(* IEC 61131-3 sources: plc_agent/plc_agent/data/rag_data/st/st_case_code, 701 files *)

(* ---- ACOSH.st ---- *)
FUNCTION ACOSH : REAL
VAR_INPUT
    X : REAL;
END_VAR
ACOSH := LN(SQRT(X * X - 1.0) + X);

(* revision history
hm		12 jan 2007	rev 1.0
	original version

hm		2. dec 2007	rev 1.1
	changed code for better performance

hm	16. mar. 2007		rev 1.2
	changed sequence of calculations to improve performance

hm	10. mar. 2009		rev 1.3
	real constants updated to new systax using dot

*)
END_FUNCTION

(* ---- ACOTH.st ---- *)
FUNCTION ACOTH : REAL
VAR_INPUT
    X : REAL;
END_VAR
ACOTH := LN((x+1.0)/(x-1.0))*0.5;

(* revision history
hm		12 jan 2007	rev 1.0
	original version

hm		5. jan 2008	rev 1.1
	improved code for better performance

hm	10. mar. 2009		rev 1.2
	real constants updated to new systax using dot

*)
END_FUNCTION

(* ---- AGDF.st ---- *)
FUNCTION AGDF : REAL
VAR_INPUT
    X : REAL;
END_VAR
AGDF := LN((1.0 + SIN(X)) / COS(X));

(* comment
the current implementation gives sufficient accuracy only up to X = 1.57 or an output > 10.
is X closer to PI/2 then the function is more and more unreliable
*)

(* revision history
hm	27. apr. 2008	rev 1.0
	original version

hm	10. mar. 2009	rev 1.1
	real constants updated to new systax using dot

*)
END_FUNCTION

(* ---- AIN.st ---- *)
FUNCTION AIN : REAL
VAR_INPUT
    in : DWORD;
    Bits : BYTE;
    sign : BYTE := 255;
    low : REAL;
    high : REAL := 10.0;
END_VAR

VAR_CONSTANT
    ff : DWORD := 16#FFFFFFFF;
END_VAR

VAR
    temp1 : DWORD;
    temp2 : DWORD;
    sx : BOOL;
END_VAR
(* extract the sign bit *)
IF sign < 32 THEN
	temp1 := SHR(in,sign);
	sx := temp1.0;
ELSE
	sx := FALSE;
END_IF;
temp1 := SHR(ff, 32-bits);
temp2 := in AND temp1;
AIN := (high - low) * DWORD_TO_REAL(temp2) / DWORD_TO_REAL(temp1) + low;
IF sx THEN AIN := -AIN; END_IF;

(* revision history
hm 18.8.2006	rev 1.1
	fixed an error with low value negative and high value 0.

hm 19.1.2007	rev 1.2
	fixed an error with sign bit.

hm	13.9.2007	rev 1.3
	changed code to avoid warning under codesys 2.8.1

hm	2. dec 2007	rev 1.4
	changed code for better performance

hm	16. mar 2008	rev 1.5
	added type conversions to avoid warnings under codesys 30
*)
END_FUNCTION

(* ---- AIR_DENSITY.st ---- *)
FUNCTION AIR_DENSITY : REAL
VAR_INPUT
    T : REAL;     // Temperature
    P : REAL;     // Pressure
    RH : REAL;    // Relative Humidity
END_VAR

VAR CONSTANT
    RL : REAL := 287.05;   // Constant value for RL
    RX : REAL := 0.003773319;  // Constant value for RX
END_VAR
AIR_DENSITY := OSCAT_BASIC.phys.PN * (1.0 - RH * SDD(T, TRUE) * RX / P) / (RL * ( T - OSCAT_BASIC.phys.T0));

(* original code used for rev 1.0

SDD := SDD(T,FALSE);
RF := RL / (1- RH*SDD/P*RX);
Air_density := P / (RF * (T-TK));

*)

(* revision history

hm	29.10.2007	rev 1.0
	original version

hm	4.12.2007		rev 1.1
	changed code for better performance

hm	18. oct. 2008	rev 1.2
	using phys constants

hm	13. mar. 2009	rev 1.3
	real constants updated to new systax using dot

*)
END_FUNCTION

(* ---- AIR_ENTHALPY.st ---- *)
FUNCTION AIR_ENTHALPY : REAL
VAR_INPUT
    T : REAL;
    RH : REAL;
END_VAR

VAR CONSTANT
    CPL : REAL := 1.00482;
    CW : REAL := 1.86;
    LH : REAL := 2500.78;
END_VAR
AIR_ENTHALPY := CPL * T + (CW * T + LH) * DEW_CON(RH,T);

(* revision history

hm	31.10.2007	rev 1.0
	original version

hm	2.11.2007		rev 1.1
	deleted unused variable RF

hm	2.12.2007		rev 1.2
	changed code for better performance
*)
END_FUNCTION

(* ---- AOUT.st ---- *)
FUNCTION AOUT : DWORD
VAR_INPUT
    in : REAL;
    Bits : BYTE;
    sign : BYTE := 255;
    low : REAL;
    high : REAL := 10.0;
END_VAR_INPUT

VAR CONSTANT
    ff : DWORD := 2#1;
END_VAR_CONSTANT

VAR
    in2 : REAL;
    sx : BOOL;
END_VAR
(* if sign bit is defined *)
IF sign < 32 THEN
	sx := sign_R(in);
	in2 := ABS(in);
ELSE
	in2 := in;
END_IF;

(* begrenze in auf die zulässigen werte *)
in2 := LIMIT(low, in2, high);

(* Berechne den Ausgangswert *)
Aout := REAL_TO_DWORD((in2 - low) / (high - low) * DWORD_TO_REAL(SHL(ff,bits) -1));
IF sx THEN Aout := SHL(ff,sign) OR Aout; END_IF;

(*
revision history

hm 18.1.2007		rev 1.1
	renamed Modul to aout.
	changed Output to 32 Bit max.
	corrected error with sign bit.

hm	13.9.2007		rev 1.2
	changed code to avoid warning under codesys 2.8.1

hm	2. dec 2007		rev 1.3
	changed code for better performance

hm	23. feb 2008	rev 1.4
	changed code for better performance
*)
END_FUNCTION

(* ---- AOUT1.st ---- *)
FUNCTION AOUT1 : DWORD
VAR_INPUT
    in : REAL;
    Bit_0 : INT; // input_constant attribute
    Bit_N : INT := 31; // input_constant attribute, initial value set
    sign : INT := 255; // input_constant attribute, initial value set
    low : REAL; // input_constant attribute
    high : REAL := 10.0; // initial value set, input_constant attribute
END_VAR

VAR CONSTANT
    ff : DWORD := 2#1; // initial value set
END_VAR

VAR
    sx : BOOL;
    in2 : REAL;
END_VAR
(* if sign bit is defined *)
IF sign < 32 THEN
	sx := SIGN_R(in);
	in2 := ABS(in);
ELSE
	in2 := in;
END_IF;

(* begrenze in auf die zulässigen werte *)
in2 := LIMIT(low, in2, high);

(* Berechne den Ausgangswert *)
AOUT1 := SHL(REAL_TO_DWORD((in2 - low) / (high - low) * DWORD_TO_REAL(SHL(ff,bit_n - Bit_0 + 1) -1)),Bit_0);
IF sx THEN AOUT1 := SHL(ff,sign) OR AOUT1; END_IF;

(* revision history
hm	23. feb 2008	rev 1.0
	original version

*)
END_FUNCTION

(* ---- ARRAY_AVG.st ---- *)
FUNCTION ARRAY_AVG : REAL
VAR_INPUT
    pt : POINTER TO ARRAY [0..32000] OF REAL;
    size : UINT;
END_VAR

VAR
    i : UINT;
    stop : UINT;
END_VAR
stop := SHR(size,2)-1;
ARRAY_AVG := pt^[0];
FOR i := 1 TO stop DO
	ARRAY_AVG := ARRAY_AVG + pt^[i];
END_FOR;
ARRAY_AVG := ARRAY_AVG / UINT_TO_REAL(stop + 1);

(* revision history
hm	2. oct 2007		rev 1.0
	original version

hm	12. dec 2007	rev 1.1
	chaged code for better performance

hm	16. mar. 2008	rev 1.2
	changed input size to uint

hm	10. mar. 2009	rev 1.3
	added type conversion for compatibility reasons
*)
END_FUNCTION

(* ---- ARRAY_GAV.st ---- *)
FUNCTION ARRAY_GAV : REAL
VAR_INPUT
    pt : POINTER TO ARRAY[0..32000] OF REAL;
    size : UINT;
END_VAR

VAR
    i : UINT;
    stop : UINT;
END_VAR
stop := SHR(size,2)-1;
ARRAY_GAV := 1.0;
FOR i := 0 TO stop DO
	IF pt^[i] > 0.0 THEN
		ARRAY_GAV := ARRAY_GAV * pt^[i];
	ELSE
		ARRAY_GAV := 0.0;
		RETURN;
	END_IF;
END_FOR;
ARRAY_GAV := SQRTN(ARRAY_GAV,UINT_TO_INT(stop)+1);

(* revision history
hm	2. apr 2008	rev 1.0
	original version

hm	10. mar. 2009	rev 1.1
	real constants updated to new systax using dot

*)
END_FUNCTION

(* ---- ARRAY_HAV.st ---- *)
FUNCTION ARRAY_HAV : REAL
VAR_INPUT
    pt    : POINTER TO ARRAY [0..32000] OF REAL;
    size  : UINT;
END_VAR

VAR
    i     : UINT;
    stop  : UINT;
END_VAR
stop := SHR(size,2)-1;
FOR i := 0 TO stop DO
	IF pt^[i] <> 0.0 THEN
		ARRAY_HAV := ARRAY_HAV + 1.0 / pt^[i];
	ELSE
		ARRAY_HAV := 0.0;
		RETURN;
	END_IF;
END_FOR;
ARRAY_HAV := UINT_TO_REAL(stop + 1) / ARRAY_HAV;

(* revision history
hm	2. apr 2008	rev 1.0
	original version

hm	10. mar. 2009	rev 1.1
	real constants updated to new systax using dot

*)
END_FUNCTION

(* ---- ARRAY_MAX.st ---- *)
FUNCTION ARRAY_MAX : REAL
VAR_INPUT
    pt : ^ARRAY[0..32000] OF REAL;
    size : UINT;
END_VAR

VAR
    i : UINT;
    stop : UINT;
END_VAR
stop := (size -SIZEOF(pt)) / SIZEOF(pt);
array_max := pt^[0];
FOR i := 1 TO stop DO
	IF pt^[i] > array_max THEN array_max := pt^[i]; END_IF;
END_FOR;

(* revision history
hm	2. oct 2006		rev 1.0
	original version

hm	16. mar. 2008	rev 1.1
	changed input size to uint
*)
END_FUNCTION

(* ---- ARRAY_MIN.st ---- *)
FUNCTION ARRAY_MIN : REAL
VAR_INPUT
    pt : POINTER TO ARRAY[0..32000] OF REAL;
    size : UINT;
END_VAR

VAR
    i : UINT;
    stop : UINT;
END_VAR
stop := (size - SIZEOF(pt)) / SIZEOF(pt);
array_min := pt^[0];
FOR i := 1 TO stop DO
	IF pt^[i] < array_min THEN array_min := pt^[i]; END_IF;
END_FOR;

(* revision history
hm		2. oct. 2006
	original version

hm		16. mar. 2008
	changed type of input size to uint

*)
END_FUNCTION

(* ---- ARRAY_SDV.st ---- *)
FUNCTION ARRAY_SDV : REAL
VAR_INPUT
    pt : POINTER TO ARRAY[0..32000] OF REAL;
    size : UINT;
END_VAR
(* standard deviation is simply the square root of the variance *)

array_sdv := SQRT(array_var(pt, size));

(* revision history
hm 	1.4.2007		rev 1.0
	function created

hm	16. mar. 2008	rev 1.1
	changed type of input size to uint

*)
END_FUNCTION

(* ---- ARRAY_SPR.st ---- *)
FUNCTION ARRAY_SPR : REAL
VAR_INPUT
    pt : ^ARRAY [0..32000] OF REAL;
    size : UINT;
END_VAR

VAR
    i : UINT;
    stop : UINT;
    array_max : REAL;
    array_min : REAL;
END_VAR
stop := (size -SIZEOF(pt)) / SIZEOF(pt);
array_min := pt^[0];
array_max := pt^[0];
FOR i := 1 TO stop DO
	IF pt^[i] > array_max THEN array_max := pt^[i];
	ELSIF pt^[i] < array_min THEN array_min := pt^[i];
	END_IF;
END_FOR;
array_spr := array_max - array_min;

(* revision history
hm 	2. oct. 2006	rev 1.0
	original version

hm	16. mar. 2008	rev 1.1
	changed type of input size to uint

*)
END_FUNCTION

(* ---- ARRAY_SUM.st ---- *)
FUNCTION ARRAY_SUM : REAL
VAR_INPUT
    pt : POINTER TO ARRAY[0..32000] OF REAL;
    size : UINT;
END_VAR_INPUT

VAR
    i : UINT;
    stop : UINT;
END_VAR
stop := (size -SIZEOF(pt)) / SIZEOF(pt);
array_sum := pt^[0];
FOR i := 1 TO stop DO
	array_sum := array_sum + pt^[i];
END_FOR;

(* revision history
hm 	2. oct. 2006	rev 1.0
	function created

hm	16. mar. 2008	rev 1.1
	changed type of input size to uint

*)
END_FUNCTION

(* ---- ARRAY_TREND.st ---- *)
FUNCTION ARRAY_TREND : REAL
VAR_INPUT
    pt : POINTER TO ARRAY[0..32000] OF REAL;
    size : UINT;
END_VAR

VAR
    i : UINT;
    stop : UINT;
    x : REAL;
    stop2 : UINT;
END_VAR
stop := SHR(size,2)-1;
stop2 := SHR(stop,1);
FOR i := 0 TO stop2 DO x := x - pt^[i]; END_FOR;
IF EVEN(UINT_TO_INT(stop)) THEN
	FOR i := stop2 TO stop DO X := X + pt^[i]; END_FOR;
ELSE
	FOR i := stop2 + 1 TO stop DO X := X + pt^[i]; END_FOR;
END_IF;
ARRAY_TREND := x / UINT_TO_REAL(stop2 + 1);

(* revision history
hm	2 oct 2007	rev 1.0
	original version

hm	12 dec 2007	rev 1.1
	changed code for better performance

hm	16. mar. 2008	rev 1.2
	changed type of input size to uint

hm	10. mar. 2009	rev 1.3
	added type conversions for compatibility reasons
*)
END_FUNCTION

(* ---- ARRAY_VAR.st ---- *)
FUNCTION ARRAY_VAR : REAL
VAR_INPUT
    pt : POINTER TO ARRAY[0..32000] OF REAL;
    size : UINT;
END_VAR

VAR
    avg : REAL;
    i : UINT;
    stop : UINT;
END_VAR
(* at first we calualte the arithmetic average of the array *)

stop := SHR(size,2)-1;
avg := pt^[0];
FOR i := 1 TO stop DO
	avg := avg + pt^[i];
END_FOR;
avg := avg / UINT_TO_REAL(stop + 1);

(* in a second run we calculate the variance of the array *)

array_var := (pt^[0] - avg) * (pt^[0] - avg);
FOR i := 1 TO stop DO
	array_var := array_var + (pt^[i] - avg) * (pt^[i] - avg);
END_FOR;
ARRAY_VAR := ARRAY_VAR / UINT_TO_REAL(stop);

(* revision history
hm 	1.4.2007	rev 1.0
	function created

hm	12.12.2007	rev 1.1
	changed code for better performance

hm	16. mar. 2008	rev 1.2
	changed type of input size to uint

hm	10. mar. 2009	rev 1.3
	added type conversions for compatibility reasons
*)
END_FUNCTION

(* ---- ASINH.st ---- *)
FUNCTION ASINH : REAL
VAR_INPUT
    X : REAL;
END_VAR
ASINH := LN(SQRT(X * X + 1.0)+X);

(* revision history
hm		12 jan 2007	rev 1.0
	original version

hm		2. dec 2007	rev 1.1
	changed code for better performance

hm		16.3. 2007		rev 1.2
	changed sequence of calculations to improve performance

hm	10. mar. 2009		rev 1.3
	real constants updated to new systax using dot

*)
END_FUNCTION

(* ---- ATAN2.st ---- *)
FUNCTION ATAN2 : REAL
VAR_INPUT
    Y : REAL;
    X : REAL;
END_VAR
IF X > 0.0 THEN
	ATAN2 := ATAN(Y/X);
ELSIF X < 0.0 THEN
	IF Y >=0.0 THEN
		ATAN2 := ATAN(Y/X) + MATH.PI;
	ELSE
		ATAN2 := ATAN(Y/X) - MATH.PI;
	END_IF;
ELSIF Y > 0.0 THEN
	ATAN2 := MATH.PI05;
ELSIF Y < 0.0 THEN
	ATAN2 := -MATH.PI05;
ELSE
	ATAN2 := 0.0;
END_IF;

(* revision history
hm	20.  apr. 2008	rev 1.0
	original version

hm	18. oct. 2008	rev 1.1
	changed to use math constants

hm	10. mar. 2009	rev 1.2
	real constants updated to new systax using dot

*)
END_FUNCTION

(* ---- ATANH.st ---- *)
FUNCTION ATANH : REAL
VAR_INPUT
    X : REAL;
END_VAR
ATANH := LN((1.0 + x)/(1.0 - x)) * 0.5;

(* revision history
hm		12 jan 2007	rev 1.0
	original version

hm		5. jan 2008	rev 1.1
	improved code for better performance

hm	10. mar. 2009		rev 1.2
	real constants updated to new systax using dot

*)
END_FUNCTION

(* ---- BAND_B.st ---- *)
FUNCTION BAND_B : BYTE
VAR_INPUT
    X : BYTE;
    B : BYTE;
END_VAR
IF X < B THEN
	BAND_B := 0;
ELSIF X > BYTE#255-B THEN
	BAND_B := 255;
ELSE
	BAND_B := X;
END_IF;

(* revision history
hm	21. nov. 2008	rev 1.0
	original version

*)
END_FUNCTION

(* ---- BASE64_DEMO.st ---- *)
FUNCTION BASE64_DEMO
VAR
    text1 : STRING(144) := '<4036.1076324381@guildenstern.zeitform.de>';
    text2 : STRING(192);
    text3 : STRING(144);
    BASE64_DECODE_STR : BASE64_DECODE_STR; (* Assuming BASE64_DECODE_STR is a previously defined type *)
    BASE64_ENCODE_STR : BASE64_ENCODE_STR; (* Assuming BASE64_ENCODE_STR is a previously defined type *)
    start : BOOL := TRUE;
    done1 : BOOL;
    done2 : BOOL;
END_VAR

END_FUNCTION

(* ---- BCDC_TO_INT.st ---- *)
FUNCTION BCDC_TO_INT : INT
VAR_INPUT
    IN : BYTE;
END_VAR
BCDC_TO_INT := (in AND 16#0F) + (SHR(in,4) * 10);

(* revision history
hm	13.12.2007	rev 1.0
	original version

hm	30.6.2008	rev 1.1
	changed name BCD_TO_INT to BCDC_TO_INT to avoid collision with util.lib

*)
END_FUNCTION

(* ---- BETA.st ---- *)
FUNCTION BETA : REAL
VAR_INPUT
    X : REAL;
    Y : REAL;
END_VAR
BETA := GAMMA(X) * GAMMA(Y) / GAMMA(x + y);

(* revision history
hm	26. oct. 2008	rev 1.0
	original version

*)
END_FUNCTION

(* ---- BFT_TO_MS.st ---- *)
FUNCTION BFT_TO_MS : REAL
VAR_INPUT
    BFT : INT;
END_VAR
BFT_TO_MS := EXPT(BFT, 1.5) * 0.836;

(* revision history
hm	12. 6. 2008		rev 1.0
	original version

*)
END_FUNCTION

(* ---- BIN_TO_BYTE.st ---- *)
FUNCTION BIN_TO_BYTE : BYTE
VAR_INPUT
    BIN : STRING(12);
END_VAR

VAR
    pt : POINTER TO BYTE;
    i : INT;
    X : BYTE;
    stop : INT;
END_VAR
pt := ADR(bin);
stop := LEN(bin);
FOR I := 1 TO stop DO
	x := pt^;
	(* calculate the value of the digit *)
	IF X = 48 THEN
		BIN_TO_BYTE := SHL(BIN_TO_BYTE,1);
	ELSIF X = 49 THEN
		BIN_TO_BYTE := SHL(BIN_TO_BYTE,1) OR 1;
	END_IF;
	pt := pt + 1;
END_FOR;

(* revision histroy
hm	18. jun. 2008	rev 1.0
	original release

hm	20. sep. 2008	rev 1.1
	changed length of input string from 20 to 12

hm	26. jul. 2009	rev 1.2
	optimized code
*)
END_FUNCTION

(* ---- BIN_TO_DWORD.st ---- *)
FUNCTION BIN_TO_DWORD : DWORD
VAR_INPUT
    BIN : STRING(40);
END_VAR

VAR
    pt : POINTER TO BYTE;
    i : INT;
    X : BYTE;
    stop : INT;
END_VAR
pt := ADR(bin);
stop := LEN(bin);
FOR I := 1 TO stop DO
	x := pt^;
	(* calculate the value of the digit *)
	IF X = 48 THEN
		BIN_TO_DWORD := SHL(BIN_TO_DWORD,1);
	ELSIF X = 49 THEN
		BIN_TO_DWORD := SHL(BIN_TO_DWORD,1) OR 1;
	END_IF;
	pt := pt + 1;
END_FOR;

(* revision histroy
hm	18. jun. 2008	rev 1.0
	original release

hm	20. sep. 2008	rev 1.1
	changed length of input dtring from 20 to 40

hm	26. jul 2009	rev 1.2
	optimized code
*)
END_FUNCTION

(* ---- BINOM.st ---- *)
FUNCTION BINOM : DINT
VAR_INPUT
    N : INT;
    K : INT;
END_VAR

VAR
    i : INT;
END_VAR
IF 2 * K > n THEN
	k := n - k;
END_IF;
IF k > n THEN
	RETURN;
ELSIF k = 0 OR k = n THEN
	BINOM := 1;
ELSIF k = 1 THEN
	BINOM := n;
ELSE
	BINOM := n;
	n := n + 1;
	FOR i := 2 TO k DO
		BINOM := BINOM * (n - i) / i;
	END_FOR;
END_IF;

(*
binomialkoeffizient(n, k)
1  wenn k = 0 return 1
2  wenn 2k > n
3      dann führe aus ergebnis \leftarrow binomialkoeffizient(n, n-k)
4  sonst führe aus ergebnis \leftarrow n
5          von i \leftarrow 2 bis k
6              führe aus ergebnis \leftarrow ergebnis \cdot (n + 1 - i)
7                        ergebnis \leftarrow ergebnis : i
8  return ergebnis
*)

(* revision history
hm	25. oct. 2008	rev 1.0
	original version

*)
END_FUNCTION

(* ---- BIT_COUNT.st ---- *)
FUNCTION BIT_COUNT : INT
VAR_INPUT
    IN : DWORD;
END_VAR
WHILE in > 0 DO
	IF in.0 THEN Bit_Count := Bit_Count + 1; END_IF;
	in := SHR(in,1);
END_WHILE;

(* revision history
5.7.2007	rev 1.0		original version

10.9.2007	rev 1.1		hm
	changed algorithm for better performace
	the execution time has reduced by a factor of 5
	deleted unused variable temp
*)
END_FUNCTION

(* ---- BIT_LOAD_B.st ---- *)
FUNCTION BIT_LOAD_B : BYTE
VAR_INPUT
    IN : BYTE;
    VAL : BOOL;
    POS : INT;
END_VAR

VAR CONSTANT
    dat : BYTE := 1;
END_VAR
IF VAL THEN
	BIT_LOAD_B := in OR SHL(dat,pos);
ELSE
	BIT_LOAD_B := in AND (NOT SHL(dat,pos));
END_IF;

(* revision history
hm	29. feb 2008	rev 1.0
	original version

hm	16. mar 2008	rev 1.1
	change input bit to val for compatibility reasons
*)
END_FUNCTION

(* ---- BIT_LOAD_B2.st ---- *)
FUNCTION BIT_LOAD_B2 : BYTE
VAR_INPUT
    I : BYTE;
    D : BOOL;
    P : INT;
    N : INT;
END_VAR
IF D THEN
	BIT_LOAD_B2 := ROL(SHR(BYTE#255, 8 - N) OR ROR(i, P), P);
ELSE
	BIT_LOAD_B2 := ROL(SHL(BYTE#255, N) AND ROR(I, P), P);
END_IF;

(* revision history
hm	18. oct. 2008	rev 1.0
	original version

*)
END_FUNCTION

(* ---- BIT_LOAD_DW.st ---- *)
FUNCTION BIT_LOAD_DW : DWORD
VAR_INPUT
    IN : DWORD;
    VAL : BOOL;
    POS : INT;
END_VAR

VAR CONSTANT
    dat : DWORD := 1;
END_VAR
IF val THEN
	BIT_LOAD_DW := in OR SHL(dat,pos);
ELSE
	BIT_LOAD_DW := in AND (NOT SHL(dat,pos));
END_IF;

(* revision history
hm	29. feb 2008	rev 1.0
	original version

hm	16. mar 2008	rev 1.1
	change input bit to val for compatibility reasons
*)
END_FUNCTION

(* ---- BIT_LOAD_DW2.st ---- *)
FUNCTION BIT_LOAD_DW2 : DWORD
VAR_INPUT
    I : DWORD;
    D : BOOL;
    P : INT;
    N : INT;
END_VAR
IF D THEN
	BIT_LOAD_DW2 := ROL(SHR(DWORD#4294967295, 32 - N) OR ROR(i, P), P);
ELSE
	BIT_LOAD_DW2 := ROL(SHL(DWORD#4294967295, N) AND ROR(I, P), P);
END_IF;

(* revision history
hm	18. oct. 2008	rev 1.0
	original version

*)
END_FUNCTION

(* ---- BIT_LOAD_W.st ---- *)
FUNCTION BIT_LOAD_W : WORD
VAR_INPUT
    IN : WORD;
    VAL : BOOL;
    POS : INT;
END_VAR

VAR_CONSTANT
    dat : WORD := 1;
END_VAR
IF val THEN
	BIT_LOAD_W := in OR SHL(dat,pos);
ELSE
	BIT_LOAD_W := in AND (NOT SHL(dat,pos));
END_IF;

(* revision history
hm	29. feb 2008	rev 1.0
	original version

hm	16. mar 2008	rev 1.1
	change input bit to val for compatibility reasons
*)
END_FUNCTION

(* ---- BIT_LOAD_W2.st ---- *)
FUNCTION BIT_LOAD_W2 : WORD
VAR_INPUT
    I : WORD;
    D : BOOL;
    P : INT;
    N : INT;
END_VAR
IF D THEN
	BIT_LOAD_W2 := ROL(SHR(WORD#65535, 16 - N) OR ROR(i, P), P);
ELSE
	BIT_LOAD_W2 := ROL(SHL(WORD#65535, N) AND ROR(I, P), P);
END_IF;

(* revision history
hm	18. oct. 2008	rev 1.0
	original version

*)
END_FUNCTION

(* ---- BIT_OF_DWORD.st ---- *)
FUNCTION BIT_OF_DWORD : BOOL
VAR_INPUT
    in : DWORD;
    N : INT;
END_VAR
BIT_OF_DWORD := (SHR(in,N) AND 16#00000001) > 0;

(* old code used before rev 1.1
temp := SHR(in,n);
Bit_of_Dword := temp.0;
*)

(* revision history
hm	4. aug. 2006	rev 1.0
	original version

hm	29. feb 2008	rev 1.1
	improved performance

hm	6. jun. 2008	rev 1.2
	changes type of input N from byte to int
*)
END_FUNCTION

(* ---- BIT_TOGGLE_B.st ---- *)
FUNCTION BIT_TOGGLE_B : BYTE
VAR_INPUT
    IN : BYTE;
    POS : INT;
END_VAR
BIT_TOGGLE_B := SHL(BYTE#1, POS) XOR IN;

(* revision history
hm	18. oct. 2008	rev 1.0
	original version

*)
END_FUNCTION

(* ---- BIT_TOGGLE_DW.st ---- *)
FUNCTION BIT_TOGGLE_DW : DWORD
VAR_INPUT
    IN : DWORD;
    POS : INT;
END_VAR
BIT_TOGGLE_DW := SHL(DWORD#1, POS) XOR IN;

(* revision history
hm	18. oct. 2008	rev 1.0
	original version

*)
END_FUNCTION

(* ---- BIT_TOGGLE_W.st ---- *)
FUNCTION BIT_TOGGLE_W : WORD
VAR_INPUT
    IN : WORD;
    POS : INT;
END_VAR
BIT_TOGGLE_W := SHL(WORD#1, POS) XOR IN;

(* revision history
hm	18. oct. 2008	rev 1.0
	original version

*)
END_FUNCTION

(* ---- BUFFER_COMP.st ---- *)
FUNCTION BUFFER_COMP : INT
VAR_INPUT
    PT1 : POINTER TO ARRAY [0..32767] OF BYTE;
    SIZE1 : INT;
    PT2 : POINTER TO ARRAY [0..32767] OF BYTE;
    SIZE2 : INT;
    START : INT;
END_VAR_INPUT

VAR
    i : INT;
    j : INT;
    end : INT;
    firstbyte : BYTE;
END_VAR
(* search for first character match *)
IF size2 <= size1 THEN
	end := size1 - size2;
	firstbyte := PT2^[0];
	FOR i := START TO end DO
		IF PT1^[i] = firstbyte THEN
			(* first character matches, now compare rest of array *)
			j := 1;
			WHILE j < size2 DO
				IF pt2^[j] <> pt1^[j+i] THEN EXIT; END_IF;
				j := j + 1;
			END_WHILE;
			(* when J > size2 a match was found return the position i in buffer1 *)
			IF j = size2 THEN
				BUFFER_COMP := i;
				RETURN;
			END_IF;
		END_IF;
	END_FOR;
END_IF;
BUFFER_COMP := -1;

(*
hm 14. nov. 2008	rev 1.0
	original version

hm	12. nov. 2009	rev 1.1
	performance increase

*)
END_FUNCTION

(* ---- BUFFER_SEARCH.st ---- *)
FUNCTION BUFFER_SEARCH : INT
VAR_INPUT
    PT : POINTER TO ARRAY[0..32767] OF BYTE;
    SIZE : INT;
    STR : STRING; // STRING_LENGTH should be replaced with actual length if known
    POS : INT;
    IGN : BOOL;
END_VAR

VAR
    ps : POINTER TO ARRAY[0..STRING_LENGTH] OF BYTE; // STRING_LENGTH should be replaced with actual length if known
    chx : BYTE;
    i : INT;
    end : INT;
    k : INT;
    lx : INT;
END_VAR
ps := ADR(STR);
lx := LEN(STR);
end := MIN(SIZE - lx, SIZE - 1);
lx := lx - 1;
FOR i := pos TO end DO
	FOR k := 0 TO lx DO
		IF IGN THEN chx := TO_UPPER(pt^[i+k]); ELSE chx := pt^[i+k]; END_IF;
		IF ps^[k] <> chx THEN EXIT; END_IF;
	END_FOR;
	IF k > lx THEN
		BUFFER_SEARCH := i;
		RETURN;
	END_IF;
END_FOR;
BUFFER_SEARCH := -1;

(* revision History

hm 5. mar. 2008	rev 1.0
	original version

hm	16. mar. 2008	rev 1.1
	chaged type of input size to uint

hm	13. may. 2008	rev 1.2
	changed type of pointer to array[1..32767]
	changed size of string to STRING_LENGTH

hm	12. nov. 2009	rev 1.3
	limit end to array size

hm	25. jan. 2011	rev 1.4
	ign = True will now ignore case
	return -1 if nothing found
*)
END_FUNCTION

(* ---- BUFFER_TO_STRING.st ---- *)
FUNCTION BUFFER_TO_STRING : string
VAR_INPUT
    PT : POINTER TO ARRAY [0..32767] OF BYTE;
    SIZE : UINT;
    START : UINT;
    STOP : UINT;
END_VAR

VAR
    ps : POINTER TO BYTE;
    i : UINT;
    stp : UINT;
    sta : UINT;
END_VAR
ps := ADR(BUFFER_TO_STRING);
IF size = 0 THEN RETURN; END_IF;
sta := MIN(start, size -1);
stp := MIN(stop, size -1);

(* check for maximum string_length *)
IF UINT_TO_INT(stp - sta + 1) >= STRING_LENGTH THEN
	stp := sta + INT_TO_UINT(STRING_LENGTH) - 1;
END_IF;

FOR i := sta TO stp DO
	ps^ := pt^[i];
	ps := ps + 1;
END_FOR;

(* terminate the string *)

ps^ := 0;

(* revision History
hm 	5. mar. 2008	rev 1.0
	original version

hm	16. mar. 2008	rev 1.1
	changed type of input size to uint

hm	13. may. 2008	rev 1.2
	changed type of pointer to array[0..32767]
	changed size of string to STRING_LENGTH

hm	12. jun. 2008	rev 1.3
	check for pointer overrun
	change input start and stop to uint
	added type conversions to avoid warnings under codesys 3.0

hm	23. mar. 2009	rev 1.4
	avoid writing to input stop

hm	12. nov. 2009 rev 1.5
	limit start and stop to size -1

*)
END_FUNCTION

(* ---- BUILDING_VERSION.st ---- *)
FUNCTION BUILDING_VERSION : DWORD
VAR_INPUT
    IN : BOOL;
END_VAR
IF in THEN
	BUILDING_VERSION := DATE_TO_DWORD(D#2011-02-3);
ELSE
	BUILDING_VERSION := 100;
END_IF;

(* revision history
hm	6. oct 2006	rev 1.0
	original version

hm	16. dec 2007	rev 1.1
	added possibility to return date and version depending on IN.

*)
END_FUNCTION

(* ---- BYTE_OF_BIT.st ---- *)
FUNCTION BYTE_OF_BIT : BYTE
VAR_INPUT
    B0 : BOOL;
    B1 : BOOL;
    B2 : BOOL;
    B3 : BOOL;
    B4 : BOOL;
    B5 : BOOL;
    B6 : BOOL;
    B7 : BOOL;
END_VAR
Byte_of_bit := SHL(SHL(SHL(SHL(SHL(SHL(SHL(BOOL_TO_BYTE(B7),1) OR BOOL_TO_BYTE(B6),1) OR BOOL_TO_BYTE(B5),1) OR BOOL_TO_BYTE(B4),1)
	OR BOOL_TO_BYTE(B3),1) OR BOOL_TO_BYTE(B2),1) OR BOOL_TO_BYTE(B1),1) OR BOOL_TO_BYTE(B0);

(* revision history

hm	4. aug 2006		rev 1.0
	original version

hm	18. feb. 2008	rev 1.1
	improved performance

*)
END_FUNCTION

(* ---- BYTE_OF_DWORD.st ---- *)
FUNCTION BYTE_OF_DWORD : BYTE
VAR_INPUT
    in : DWORD;
    N : BYTE;
END_VAR
BYTE_OF_DWORD := DWORD_TO_BYTE(SHR(in,SHL(n,3)));

(* revision history
hm	17. jan 2007	rev 1.0
	original version

hm	2. jan 2008		rev 1.1
	improved performance

hm	30. oct. 2008	rev 1.2
	improved performance
*)
END_FUNCTION

(* ---- BYTE_TO_GRAY.st ---- *)
FUNCTION BYTE_TO_GRAY : BYTE
VAR_INPUT
    IN : BYTE;
END_VAR
BYTE_TO_GRAY := IN XOR SHR(IN,1);

(* revision history
hm	9. nov. 2009	rev 1.0
	original version

*)
END_FUNCTION

(* ---- BYTE_TO_RANGE.st ---- *)
FUNCTION BYTE_TO_RANGE : REAL
VAR_INPUT
    X : BYTE;
    low : REAL;
    high : REAL;
END_VAR
BYTE_TO_RANGE := (high - low) * X / 255.0 + low;

(* revision history
hm	9. jan 2008		rev 1.0
	original version

*)
END_FUNCTION

(* ---- BYTE_TO_STRB.st ---- *)
FUNCTION BYTE_TO_STRB : string
VAR_INPUT
    IN : BYTE;
END_VAR

VAR
    i : INT;
    pt : POINTER TO BYTE;
END_VAR
(* pointer für die ausgabe ermitteln *)
pt := ADR(BYTE_TO_STRB);
(* die 8 ausgabecharacter ermitteln und schreiben *)
FOR i := 1 TO 8 DO
	pt^ := BOOL_TO_BYTE(in.7) + 48;
	in := SHL(in,1);
	pt := pt + 1;
END_FOR;

(* der ausgabestring muss noch mit 0 abgeschlossen werden *)
pt^ := 0;

(* code before rev 1.1
FOR i := 1 TO 8 DO
	IF in.0 = 0 THEN temp := CONCAT('0', temp); ELSE temp := CONCAT('1', temp); END_IF;
	in := SHR(in, 1);
END_FOR;
BYTE_TO_STRB := temp;
*)

(* revision history

hm		9.6.2007	rev 1.0
	original version

hm	15. dec 2007	rev 1.1
	inprooved code for higher performance

hm	29. mar. 2008	rev 1.2
	changed STRING to STRING(8)

hm	20. jun. 2008	rev 1.3
	performance improvement

*)
END_FUNCTION

(* ---- BYTE_TO_STRH.st ---- *)
FUNCTION BYTE_TO_STRH : string
VAR_INPUT
    IN : BYTE; // Input variable
END_VAR

VAR
    temp : BYTE; // Local variable
    PT : POINTER TO BYTE; // Pointer to a BYTE
END_VAR
(* read pointer to output string *)
PT := ADR(BYTE_TO_STRH);
(* calculate high order hex value *)
temp := SHR(in,4);
(* convert value to hex character *)
IF temp <= 9 THEN temp := temp + 48; ELSE temp := temp + 55; END_IF;
(* write friat character to output string *)
PT^ := temp;
(* calculate low order hex value *)
temp := in AND 2#00001111;
IF temp <= 9 THEN temp := temp + 48; ELSE temp := temp + 55; END_IF;
(* increment pointer and wirte low order character *)
pt := pt + 1;
pt^ := temp;
(* set pointer at the end of the output string and close the string with 0 *)
pt := pt + 1;
pt^:= 0;

(* code before rev 1.2
FOR i := 1 TO 2 DO
	X := in AND 2#1111;
	IF X <= 9 THEN X := X + 48; ELSE X := X + 55; END_IF;
	Cx := CHR(X);
	temp := CONCAT(Cx, temp);
	in := SHR(in,4);
END_FOR;
BYTE_TO_STRH := temp;
*)

(* revision history

hm	9.6.2007		rev 1.0
	original version

hm	11.9.2007		rev 1.1
	changed coding for compatibility with twincat, under twincat concat cannot have a function as argument.

hm	15 dec 2007		REV 1.2
	changed code for higher performance

hm	29. mar. 2008	rev 1.3
	changed STRING to STRING(2)
*)
END_FUNCTION

(* ---- C_TO_F.st ---- *)
FUNCTION C_TO_F : REAL
VAR_INPUT
    celsius : REAL;
END_VAR
C_TO_F := celsius * 1.8 + 32.0;

(* revision history

hm	4. aug. 2006	rev 1.0
	original version

hm	11. mar. 2009	rev 1.1
	real constants updated to new systax using dot

*)
END_FUNCTION

(* ---- C_TO_K.st ---- *)
FUNCTION C_TO_K : REAL
VAR_INPUT
    Celsius : REAL;
END_VAR
C_TO_K := Celsius - phys.T0;

(* revision history

hm	4. aug 2006	rev 1.0
	original version

hm	19. aug 2009	rev 1.1
	fixed calculation error

*)
END_FUNCTION

(* ---- CABS.st ---- *)
FUNCTION CABS : REAL
VAR_INPUT
    X : COMPLEX;
END_VAR
CABS := HYPOT(x.re, x.im);

(* revision history
hm	21. feb 2008	rev 1.0
	original version

*)
END_FUNCTION

(* ---- CACOS.st ---- *)
FUNCTION CACOS : complex
VAR_INPUT
    X : COMPLEX;
END_VAR

VAR
    Y : COMPLEX;
END_VAR
y := CACOSH(x);
CACOS.re := y.im;
CACOS.im := -y.re;

(* revision history
hm	21. feb 2008	rev 1.0
	original version

*)
END_FUNCTION

(* ---- CACOSH.st ---- *)
FUNCTION CACOSH : complex
VAR_INPUT
    X : COMPLEX; // Input variable
END_VAR

VAR
    Y : COMPLEX; // Local variable
END_VAR
y.re := (X.re - X.im)*(X.re + X.im) - 1.0;
y.im := 2.0 * X.re * X.im;
y    := CSQRT(y);
y.re := y.re + x.re;
y.im := y.im + x.im;
CACOSH  := CLOG(y);

(* revision history
hm	21. feb 2008	rev 1.0
	original version

*)
END_FUNCTION

(* ---- CADD.st ---- *)
FUNCTION CADD : complex
VAR_INPUT
    X : complex;
    Y : complex;
END_VAR
CADD.re := x.re + y.re;
CADD.im := x.im + y.im;

(* revision history
hm	21. feb 2008	rev 1.0
	original version

*)
END_FUNCTION

(* ---- CAPITALIZE.st ---- *)
FUNCTION CAPITALIZE : string
VAR_INPUT
    str : STRING(STRING_LENGTH);
END_VAR

VAR
    PT : POINTER TO BYTE;
    pos : INT;
    L : INT;
    first : BOOL := TRUE;
END_VAR
PT := ADR(CAPITALIZE);
CAPITALIZE := str;
L := LEN(str);
FOR pos := 1 TO l DO
	IF first THEN pt^ := TO_UPPER(pt^);	END_IF;
	(* remember in first if the next char needs to capitalized *)
	first := pt^= 32;
	PT := pt + 1;
END_FOR;

(* revision histroy
hm		4. mar 2008	rev 1.0
	original release

hm	29. mar. 2008	rev 1.1
	changed STRING to STRING(STRING_LENGTH)

hm	20. jun. 2008	rev 1.2
	improved performance

*)
END_FUNCTION

(* ---- CARG.st ---- *)
FUNCTION CARG : REAL
VAR_INPUT
    X: COMPLEX;
END_VAR
CARG := ATAN2(X.im, X.re);

(* revision history
hm	21. feb. 2008	rev 1.0
	original version

hm	20. apr. 2008	rev 1.1
	use ATAN2 instead of ATAN
*)
END_FUNCTION

(* ---- CASIN.st ---- *)
FUNCTION CASIN : complex
VAR_INPUT
    X : complex; (* Input variable of type complex *)
END_VAR

VAR
    Y : complex; (* Local variable of type complex *)
END_VAR
y.re := -x.im;
y.im := x.re;
y := CASINH(y);
CASIN.re := y.im;
CASIN.im := -y.re;

(* revision history
hm	21. feb 2008	rev 1.0
	original version

*)
END_FUNCTION

(* ---- CASINH.st ---- *)
FUNCTION CASINH : complex
VAR_INPUT
    X : complex;
END_VAR_INPUT

VAR
    Y : complex;
END_VAR
y.re := (X.re - X.im)*(X.re + X.im) + 1.0;
y.im := 2.0 * X.re * X.im;
y    := CSQRT(y);
y.re := y.re + x.re;
y.im := y.im + x.im;
CASINH  := CLOG(y);

(* revision history
hm	21. feb 2008	rev 1.0
	original version

*)
END_FUNCTION

(* ---- CATAN.st ---- *)
FUNCTION CATAN : complex
VAR_INPUT
    X : complex; (* Input variable of type complex *)
END_VAR

VAR
    r2 : REAL;   (* Local variable of type REAL *)
    num : REAL;  (* Local variable of type REAL *)
    den : REAL;  (* Local variable of type REAL *)
END_VAR
r2 := x.re * x.re;
den := 1.0 - r2 - x.im * x.im;
CATAN.re := 0.5 * ATAN(2.0 * x.re / den);
num := x.im + 1.0;
num := r2 + num * num;
den := x.im - 1.0;
den := r2 + den * den;
CATAN.im := 0.25 * (LN(num)-LN(den));

(* revision history
hm	21. feb 2008	rev 1.0
	original version

*)
END_FUNCTION

(* ---- CATANH.st ---- *)
FUNCTION CATANH : complex
VAR_INPUT
    X : complex;
END_VAR

VAR
    i2 : REAL;
    num : REAL;
    den : REAL;
END_VAR
i2 := x.im * x.im;
num := 1.0 + x.re;
num := i2 + num * num;
den := 1.0 - x.re;
den := i2 + den * den;
CATANH.re := 0.25 * (LN(num) - LN(den));
den := 1 - x.re * x.re - i2;
CATANH.im := 0.5 * ATAN(2.0 * x.im / den);

(* revision history
hm	21. feb 2008	rev 1.0
	original version

*)
END_FUNCTION

(* ---- CAUCHY.st ---- *)
FUNCTION CAUCHY : REAL
VAR_INPUT
    X : REAL;
    T : REAL;
    U : REAL;
END_VAR

VAR
    tmp : REAL;
END_VAR
tmp := x - t;
CAUCHY := math.PI_INV * U / (U*U + tmp*tmp);

(* revision hisdtory
hm	26. oct. 2008	rev 1.0
	original version

*)
END_FUNCTION

(* ---- CAUCHYCD.st ---- *)
FUNCTION CAUCHYCD : REAL
VAR_INPUT
    X : REAL;
    T : REAL;
    U : REAL;
END_VAR
CAUCHYCD := 0.5 + math.PI_INV * ATAN((X - T) / U);

(* revision hisdtory
hm	26. oct. 2008	rev 1.0
	original version

*)
END_FUNCTION

(* ---- CCON.st ---- *)
FUNCTION CCON : complex
VAR_INPUT
    X : COMPLEX;
END_VAR
CCON.re := x.re;
CCON.im := -x.im;

(* revision history
hm	21. feb 2008	rev 1.0
	original version

*)
END_FUNCTION

(* ---- CCOS.st ---- *)
FUNCTION CCOS : complex
VAR_INPUT
    X : COMPLEX;
END_VAR
CCOS := CCOSH(CSET(-X.im, X.re));

(* revision history
hm	21. feb 2008	rev 1.0
	original version

*)
END_FUNCTION

(* ---- CCOSH.st ---- *)
FUNCTION CCOSH : complex
VAR_INPUT
    X : COMPLEX;
END_VAR
CCOSH.re := cosH(x.re) * COS(x.im);
CCOSH.im := sinH(x.re) * SIN(x.im);

(* revision history
hm	21. feb 2008	rev 1.0
	original version

*)
END_FUNCTION

(* ---- CDIV.st ---- *)
FUNCTION CDIV : complex
VAR_INPUT
    X : complex;
    Y : complex;
END_VAR

VAR
    Temp : REAL;
END_VAR
temp := Y.re * Y.re + Y.im * Y.im;
CDIV.re := (X.re * Y.re + X.im * Y.im) / temp;
CDIV.im := (X.im * Y.re - X.re * Y.im) / temp;

(* revision history
hm	21. feb 2008	rev 1.0
	original version

*)
END_FUNCTION

(* ---- CEIL.st ---- *)
FUNCTION CEIL : INT
VAR_INPUT
    X : REAL;
END_VAR
CEIL := REAL_TO_INT(x);
IF CEIL < X THEN
	CEIL := CEIL + 1;
END_IF;

(* revision history
hm	7. feb. 2007	rev 1.0
	original version

hm	21. mar. 2008	rev 1.1
	use REAL_TO_INT instead of trunc for compatibility reasons

*)
END_FUNCTION

(* ---- CEIL2.st ---- *)
FUNCTION CEIL2 : DINT
VAR_INPUT
    X: REAL;
END_VAR
CEIL2 := REAL_TO_DINT(X);
IF DINT_TO_REAL(CEIL2) < X THEN
	CEIL2 := CEIL2 + 1;
END_IF;

(* revision history
hm	21. mar. 2008	rev 1.0
	original version

hm	4. apr. 2008	rev 1.1
	added type conversion to avoid warnings under codesys 3.0

hm	30. jun. 2008	rev 1.2
	added type conversion to avoid warnings under codesys 3.0

hm	10. mar. 2009	rev 1.3
	use correct statement real_to_DINT

*)
END_FUNCTION

(* ---- CEXP.st ---- *)
FUNCTION CEXP : complex
VAR_INPUT
        X : COMPLEX;
    END_VAR

    VAR
        Temp : REAL;
    END_VAR
temp := EXP(X.re);
CEXP.re := temp * COS(X.im);
CEXP.im := temp * SIN(X.im);

(* revision history
hm	21. feb 2008	rev 1.0
	original version

*)
END_FUNCTION

(* ---- CHARCODE.st ---- *)
FUNCTION CHARCODE : BYTE
VAR_INPUT
    STR : STRING[10];
END_VAR

VAR
    found : STRING[1];
    search : STRING[10];
    pos : INT;
    i : INT;
END_VAR
IF LEN(str) = 1 THEN
	CHARCODE := CODE(STR, 1);
ELSIF str <> '' THEN
	(* construct search string *)
	search := CONCAT('&', str);
	search := CONCAT(search, ';');
	WHILE pos = 0 AND (i < 4) DO
		i := i + 1;
		pos := FIND(setup.CHARNAMES[i], search);
	END_WHILE;
	found := MID(setup.CHARNAMES[i], 1, pos - 1);
	CHARCODE := CODE(found, 1);
END_IF;

(* revision history
hm	13. may. 2008	rev 1.0
	original version

hm	19. oct. 2008	rev 1.1
	changed setup constants

hm	24. oct. 2008	rev 1.2
	optimized code
*)
END_FUNCTION

(* ---- CHARNAME.st ---- *)
FUNCTION CHARNAME : string
VAR_INPUT
    C : BYTE;
END_VAR

VAR
    pos : INT;
    i : INT;
END_VAR
IF C <> 0 THEN
	(* construct search string from code followed by $ sign, also clear charname string*)
	CHARNAME := CHR_TO_STRING(C);
	CHARNAME := CONCAT(CHARNAME,'&');
	CHARNAME := CONCAT(';', CHARNAME);
	WHILE pos = 0 AND (i < 4) DO
		i := i + 1;
		pos := FIND(setup.CHARNAMES[i], CHARNAME);
	END_WHILE;
	IF pos > 0 THEN
		CHARNAME := MID(setup.CHARNAMES[i], 10, pos + 3);
		(* search for end of name and truncate *)
		pos := FIND(CHARNAME, ';');
		CHARNAME := LEFT(CHARNAME,pos - 1);
	ELSE
		CHARNAME := CHR_TO_STRING(C);
	END_IF;
ELSE
	CHARNAME := '';
END_IF;

(* revision history
hm	13. may. 2008	rev 1.0
	original version

hm	16. jun. 2008	rev 1.1
	changed nested call of concat for better compatibility

hm	19. oct. 2008	rev 1.2
	changes setup constants

hm	24. oct. 2008	rev 1.3
	new code for high performance

hm	17. dec. 2008	rev 1.4
	changed function chr to chr_to_string
*)
END_FUNCTION

(* ---- CHECK_PARITY.st ---- *)
FUNCTION CHECK_PARITY : BOOL
VAR_INPUT
    in : DWORD;
    p : BOOL;
END_VAR
CHECK_PARITY := NOT p;
WHILE in > 0 DO
	CHECK_PARITY := CHECK_PARITY XOR in.0 XOR in.1 XOR in.2 XOR in.3;
	in := SHR(in,4);
END_WHILE;

(* code before rev 1.2
WHILE in > 0 DO
	IF in.0 THEN cnt := cnt + 1; END_IF;
	in := SHR(in,1);
END_WHILE;
check_parity := even(cnt) XOR P;
*)

(* revision history

rev 1.0 HM  1.oct.2006

rev 1.1 hm	10.sep.2007
	changed algorithm to improove performance

rev 1.2	hm	8 dec 2007
	changed algorithm to improove performance

rev 1.3 hm	18. feb 2008
	changed algorithm to improove performance
*)
END_FUNCTION

(* ---- CHK_REAL.st ---- *)
FUNCTION CHK_REAL : BYTE
VAR_INPUT
    X : REAL;
END_VAR

VAR
    pt : POINTER TO DWORD;
    tmp : DWORD;
END_VAR
pt := ADR(X);				(* move real to dword, real_to_dword does not work becasze it treats dword as a number on many systems *)
tmp := ROL(pt^,1);			(* rotate left foir easy checking, sign will be at lease significant digit *)
IF tmp < 16#FF000000 THEN
	CHK_REAL := 16#00;		(* normalized and denormalized numbers *)
ELSIF tmp = 16#FF000000 THEN
	CHK_REAL := 16#20;		(* X is +infinity see IEEE754 *)
ELSIF tmp = 16#FF000001 THEN
	CHK_REAL := 16#40;		(* X is -infinity see IEEE754 *)
ELSE
	CHK_REAL := 16#80;		(* X is NAN see IEEE754 *)
END_IF;

(* revision history
hm	 20. jan. 2011	rev 1.0
	original version

*)
END_FUNCTION

(* ---- CHR_TO_STRING.st ---- *)
FUNCTION CHR_TO_STRING : string
VAR_INPUT
    C : BYTE;
END_VAR

VAR
    PT : POINTER TO BYTE;
END_VAR
PT := ADR(CHR_TO_STRING);
PT^ := C;
pt := pt + 1;
pt^ := 0;

(* revision history
hm	16 jan 2007		rev 1.0
	original version

hm	4. feb. 2008	rev 1.1
	return string would not be terminated properly

hm	29. mar. 2008	rev 1.2
	changed STRING to STRING(1)

hm	17. dec. 2008	rev 1.3
	changed name of function from chr to chr_to_string
*)
END_FUNCTION

(* ---- CINV.st ---- *)
FUNCTION CINV : complex
VAR_INPUT
    X : COMPLEX; // Input variable of type complex
END_VAR

VAR
    temp : REAL; // Local variable of type REAL
END_VAR
temp := X.re * X.re + X.im * X.im;
CINV.re := X.re / temp;
CINV.im := -X.im / temp;

(* revision history
hm	21. feb 2008	rev 1.0
	original version

*)
END_FUNCTION

(* ---- CIRCLE_A.st ---- *)
FUNCTION CIRCLE_A : REAL
VAR_INPUT
    rx : REAL;
    ax : REAL;
END_VAR
circle_A := Rx * RX * 8.726646E-3 * Ax;

(* revision histroy
hm	16. oct 2007	rev 1.0
	original version

hm	4. dec 2007		rev 1.1
	changed code for better performance

hm	22. feb 2008	rev 1.2
	improved performance
*)
END_FUNCTION

(* ---- CIRCLE_C.st ---- *)
FUNCTION CIRCLE_C : REAL
VAR_INPUT
    Rx : REAL;
    Ax : REAL;
END_VAR
circle_C := 1.7453293E-2 * Rx * Ax;

(* revision histroy
hm	16. oct 2007	rev 1.0
	original version

hm	22. feb 2008	rev 1.1
	improved performance
*)
END_FUNCTION

(* ---- CIRCLE_SEG.st ---- *)
FUNCTION CIRCLE_SEG : REAL
VAR_INPUT
    RX : REAL;
    HX : REAL;
END_VAR
IF RX > 0.0 THEN
	CIRCLE_SEG := 2.0 * ACOS(1.0 - LIMIT(0.0, HX / RX, 2.0));
	CIRCLE_SEG := (CIRCLE_SEG - SIN(CIRCLE_SEG)) *RX * RX / 2.0;
END_IF;

(* revision histroy
hm	10. mar 2010	rev 1.0
	original version

*)
END_FUNCTION

(* ---- CLEAN.st ---- *)
FUNCTION CLEAN : string
VAR_INPUT
    IN : STRING[STRING_LENGTH];
    CX : STRING[80];
END_VAR

VAR
    pos : INT := 1;
    stop : INT;
END_VAR
(* copy input string *)
CLEAN := IN;
stop := LEN(in);
WHILE pos <= stop DO
	IF FIND(cx, MID(CLEAN, 1, pos)) > 0 THEN
		(* charcter found skip to next one *)
		pos := pos + 1;
	ELSE
		(* wrong chracter needs to be deleted *)
		CLEAN := DELETE(CLEAN, 1, pos);
		stop := stop - 1;	(* the string is one character shorter now *)
	END_IF;
END_WHILE;

(* revision history

hm		18. jun. 2008	rev 1.0
	original version

*)
END_FUNCTION

(* ---- CLOG.st ---- *)
FUNCTION CLOG : complex
VAR_INPUT
    X : COMPLEX; // Derived type 'complex'
END_VAR
CLOG.re := LN(HYPOT(X.re, X.im));
CLOG.im := ATAN2(X.im, X.re);

(* revision history
hm	21. feb 2008	rev 1.0
	original version

hm	20. apr. 2008	rev 1.1
	use ATAN2 instead of ATAN
*)
END_FUNCTION

(* ---- CMP.st ---- *)
FUNCTION CMP : BOOL
VAR_INPUT
    X : REAL;
    Y : REAL;
    N : INT;
END_VAR

VAR
    tmp : REAL;
END_VAR
tmp := ABS(x);
IF tmp > 0.0 THEN
	tmp := EXP10(INT_TO_REAL(FLOOR(LOG(tmp))-N+1));
ELSE
	tmp := EXP10(tmp);
END_IF;
CMP := ABS(X - Y) < tmp;

(* revision history
hm	12. mar. 2008	rev 1.0
	original version

hm	10. mar. 2009	rev 1.1
	added type conversion for compatibility reasons
*)
END_FUNCTION

(* ---- CMUL.st ---- *)
FUNCTION CMUL : complex
VAR_INPUT
    X : COMPLEX;
    Y : COMPLEX;
END_VAR
CMUL.re := X.re * Y.re - X.im * Y.im;
CMUL.im := X.re * Y.im + X.im * Y.re;

(* revision history
hm	21. feb 2008	rev 1.0
	original version

*)
END_FUNCTION

(* ---- CODE.st ---- *)
FUNCTION CODE : BYTE
VAR_INPUT
    STR : STRING[STRING_LENGTH];
    POS : INT;
END_VAR

VAR
    PT : POINTER TO BYTE;
END_VAR
IF pos < 1 OR pos > LEN(str) THEN
	CODE := 0;
	RETURN;
ELSE
	PT := ADR(STR) + INT_TO_DWORD(pos - 1);
	CODE := pt^;
END_IF;

(* revision history
hm	9. mar. 2008	rev 1.0
	original version

hm	29. mar. 2008	rev 1.1
	changed STRING to STRING(STRING_LENGTH)
*)
END_FUNCTION

(* ---- CONE_V.st ---- *)
FUNCTION CONE_V : REAL
VAR_INPUT
    rx : REAL;
    hx : REAL;
END_VAR
cone_V := 1.047197551 * RX * RX * hx;

(* revision histroy
hm	17. oct 2007	rev 1.0
	original version

hm	4. dec 2007		rev 1.1
	changed code for better performance

hm	22. feb 2008	rev 1.2
	changed code for better performance
*)
END_FUNCTION

(* ---- COSH.st ---- *)
FUNCTION COSH : REAL
VAR_INPUT
    X : REAL;
END_VAR

VAR
    t : REAL;
END_VAR
T := EXP(X);
COSH := (1.0 / T + T) * 0.5;

(* revision histroy
hm	12.1.2007	rev 1.0
	original version

hm	1.12.2007	rev 1.1
	changed code to improve performance

hm	5. jan 2008	rev 1.2
	further performance improvement

hm	10. mar. 2009	rev 1.3
	real constants updated to new systax using dot
*)
END_FUNCTION

(* ---- COTH.st ---- *)
FUNCTION COTH : REAL
VAR_INPUT
    X : REAL;
END_VAR
IF X > 20.0 THEN
	COTH :=1.0;
ELSIF X < -20.0 THEN
	COTH := -1.0;
ELSE
	COTH := 1.0 + 2.0 / (EXP(X * 2.0) - 1.0);
END_IF;

(* revision histroy
hm		12.1.2007	rev 1.0
	original version

hm	1.12.2007		rev 1.1
	changed code to improve performance

hm	8. jan 2008	rev 1.2
	further improvement in performance

hm	10. mar 2008	rev 1.3
	extended range of valid inputs to +/- INV
	changed formula for better accuracy

hm	10. mar. 2009	rev 1.4
	real constants updated to new systax using dot
*)
END_FUNCTION

(* ---- COUNT_CHAR.st ---- *)
FUNCTION COUNT_CHAR : INT
VAR_INPUT
    str : STRING[STRING_LENGTH];  // Input variable of type STRING with the specified length
    chr : BYTE;                    // Input variable of type BYTE
END_VAR

VAR
    l : INT;                       // Local variable of type INT
    pt : POINTER TO BYTE;          // Local variable that is a pointer to BYTE
    pos : INT;                     // Local variable of type INT
END_VAR
PT := ADR(str);
l := LEN(str);
COUNT_CHAR := 0;
FOR pos := 1 TO l DO
	IF pt^ = CHR THEN COUNT_CHAR := COUNT_CHAR + 1; END_IF;
    PT := PT + 1;
END_FOR;

(* revision history
hm	29. feb 2008	rev 1.0
	original version

hm	29. mar. 2008	rev 1.1
	changed STRING to STRING(STRING_LENGTH)
*)
END_FUNCTION

(* ---- COUNT_SUBSTRING.st ---- *)
FUNCTION COUNT_SUBSTRING : INT
VAR_INPUT
    SEARCH: STRING;
    STR: STRING;
END_VAR

VAR
    pos: INT;
    size: INT;
END_VAR
COUNT_SUBSTRING := 0;
size := LEN(SEARCH);
REPEAT
   pos := FIND(STR,SEARCH);
   IF pos > 0 THEN
      STR := REPLACE(STR, '', size,pos);
      COUNT_SUBSTRING := COUNT_SUBSTRING + 1;
   END_IF;
UNTIL pos = 0
END_REPEAT;

(* revision history
ks	20. jan. 2011	rev 1.0
	original version

*)
END_FUNCTION

(* ---- CPOL.st ---- *)
FUNCTION CPOL : complex
VAR_INPUT
    L: REAL;
    A: REAL;
END_VAR
CPOL.re := L * COS(A);
CPOL.im := L * SIN(A);

(* revision history
hm	21. feb 2008	rev 1.0
	original version

*)
END_FUNCTION

(* ---- CPOW.st ---- *)
FUNCTION CPOW : complex
VAR_INPUT
    X : Complex;
    Y : Complex;
END_VAR
CPOW := CEXP(CMUL(Y,CLOG(X)));

(* revision history
hm	21. feb 2008	rev 1.0
	original version

*)
END_FUNCTION

(* ---- CRC_GEN.st ---- *)
FUNCTION CRC_GEN : DWORD
VAR_INPUT
    PT : POINTER TO ARRAY[0..32000] OF BYTE;
    SIZE : INT;
    PL : INT;
    PN : DWORD;
    INIT : DWORD;
    REV_IN : BOOL;
    REV_OUT : BOOL;
    XOR_OUT : DWORD;
END_VAR

VAR
    pos : INT;
    shift : INT;
    dx : BYTE;
    bits : INT;
END_VAR
(* align polygon *)
shift := 32 - PL;
PN := SHL(PN, shift);

(* load first 4 bytes into register minimum message size is 4 bytes
	for smaller messages fill with 0#s at the beginning*)
FOR pos := 0 TO 3 DO
	IF REV_IN THEN CRC_GEN := SHL(CRC_GEN, 8) OR REVERSE(PT^[pos]); ELSE CRC_GEN := SHL(CRC_GEN, 8) OR PT^[pos]; END_IF;
END_FOR;
pos := 4;

(* xor with init value *)
CRC_GEN := CRC_GEN XOR SHL(init, shift);

(* calculate CRC for each byte *)
WHILE pos < size DO
	IF REV_IN THEN DX := REVERSE(PT^[pos]); ELSE DX := PT^[pos]; END_IF;
	pos := pos + 1;
	(* crc calculation for one byte *)
	FOR bits := 0 TO 7 DO
		IF CRC_GEN.31 THEN
			CRC_GEN := (SHL(CRC_GEN, 1) OR BOOL_TO_DWORD(DX.7)) XOR PN;
		ELSE
			CRC_GEN := SHL(CRC_GEN, 1) OR BOOL_TO_DWORD(DX.7);
		END_IF;
		dx := SHL(dx, 1);
	END_FOR;
END_WHILE;

(* all bytes are processed, need to finish the registers 32 bits *)
FOR bits := 0 TO 31 DO
	IF CRC_GEN.31 THEN
		CRC_GEN := (SHL(CRC_GEN, 1) ) XOR PN;
	ELSE
		CRC_GEN := SHL(CRC_GEN, 1);
	END_IF;
END_FOR;

(* final XOR *)
CRC_GEN := SHR(CRC_GEN, shift) XOR XOR_OUT;

(* reverse the crc_out put if necessary *)
IF REV_OUT THEN CRC_GEN := REFLECT(CRC_GEN, PL); END_IF;

(* suggested optimization by deninis klopke
die betreffs genannte Funktion kann folgendermaßen optimiert werden:
In Zeilen 33 und 35 des Implementierungsteils kann jeweils der Teil „OR BOOL_TO_DWORD(DX.7)“ entfallen, da nach 8maligem Linksshift von „DX“ in Zeile 26 der Wert von DX = BYTE#0 ist. Eine weitere Veroderung mit diesem Wert hat keine Auswirkungen auf das Ergebnis mehr.
*)

(* typical crc polynoms

CRC-4-ITU 			x4 + x + 1 					(ITU G.704, p. 12) 	0x3 or 0xC (0x9)
CRC-5-ITU 			x5 + x4 + x2 + 1 			(ITU G.704, p. 9) 	0x15 or 0x15 (0x0B) Bluetooth
CRC-5-USB 			x5 + x2 + 1 				(use: USB token packets) 	0x05 or 0x14 (0x9)
CRC-6-ITU 			x6 + x + 1 					(ITU G.704, p. 3) 	0x03 or 0x30 (0x21)
CRC-7 				x7 + x3 + 1 				(use: telecom systems, MMC) 	0x09 or 0x48 (0x11)
CRC-8-ATM 			x8 + x2 + x + 1 				(use: ATM HEC) 	0x07 or 0xE0 (0xC1)
CRC-8-CCITT 		x8 + x7 + x3 + x2 + 1 		(use: 1-Wire bus) 	0x8D or 0xB1 (0x63)
CRC-8-Dallas/Maxim 	x8 + x5 + x4 + 1 			(use: 1-Wire bus) 	0x31 or 0x8C (0x19)
CRC-8 				x8 + x7 + x6 + x4 + x2 + 1 	0xD5 or 0xAB (0x57)
CRC-8-SAE J1850 	x8 + x4 + x3 + x2 + 1 		0x1D or 0xB8
CRC-10 				x10 + x9 + x5 + x4 + x + 1 	0x233 or 0x331 (0x263)
CRC-12 				x12 + x11 + x3 + x2 + x + 1 (use: telecom systems) 	0x80F or 0xF01 (0xE03)
CRC-15-CAN 			x15 + x14 + x10 + x8 + x7 + x4 + x3 + 1 	0x4599 or 0x4CD1 (0x19A3)
CRC-16-Fletcher 	Not a CRC; see Fletcher's checksum 	Used in Adler-32 A & B CRCs
CRC-16-CCITT 	x16 + x12 + x5 + 1 (XMODEM,X.25, V.41, Bluetooth, PPP, IrDA; known as "CRC-CCITT") 	0x1021 or 0x8408 (0x0811)
CRC-16-IBM 	x16 + x15 + x2 + 1 (USB, many others; also known as "CRC-16") 	0x8005 or 0xA001 (0x4003)
CRC-24-Radix-64 	x24 + x23 + x18 + x17 + x14 + x11 + x10 + x7 + x6 + x5 + x4 + x3 + x + 1 	0x864CFB or 0xDF3261 (0xBE64C3)
CRC-32-Adler 	Not a CRC; see Adler-32 	See Adler-32
CRC-32-MPEG2 	x32 + x26 + x23 + x22 + x16 + x12 + x11 + x10 + x8 + x7 + x5 + x4 + x2 + x + 1 	0x04C11DB7 or 0xEDB88320 (0xDB710641) Also used in IEEE 802.3
CRC-32-IEEE 802.3 	x32 + x26 + x23 + x22 + x16 + x12 + x11 + x10 + x8 + x7 + x5 + x4 + x2 + x + 1 (V.42) 	0x04C11DB7 or 0xEDB88320 (0xDB710641)
CRC-32C (Castagnoli) 	x32 + x28 + x27 + x26 + x25 + x23 + x22 + x20 + x19 + x18 + x14 + x13 + x11 + x10 + x9 + x8 + x6 + 1 	0x1EDC6F41 or 0x82F63B78 (0x05EC76F1)
CRC-64-ISO 	x64 + x4 + x3 + x + 1 (use: ISO 3309) 	0x000000000000001B or 0xD800000000000000 (0xB000000000000001)
CRC-64-ECMA-182 	x64 + x62 + x57 + x55 + x54 + x53 + x52 + x47 + x46 + x45 + x40 + x39 + x38 + x37 + x35 + x33 + x32 + x31 + x29 + x27 + x24 + x23 + x22 + x21 + x19 + x17 + x13 + x12 + x10 + x9 + x7 + x4 + x + 1
(as described in ECMA-182 p.63) 	0x42F0E1EBA9EA3693 or 0xC96C5795D7870F42 (0x92D8AF2BAF0E1E85)
*)

(* revision history

hm	9.6.2007		rev 1.0
	original version

hm	11.9.2007		rev 1.1
	deleted unused variable i

hm	9. oct 2007 	rev 1.2
	added init code for crc and xor_out
	added refelct in and reflect_out (rev_in und Rev_out)

hm	2. jan 2008	rev 1.3
	small changes for performance improvements

hm	16. mar. 2008	rev 1.4
	changed type of input size to uint

hm	10. mar. 2009	rev 1.5
	removed nested comments

hm	16. jan. 2011	rev 2.0
	new version

dk 3. feb 2021		rev 2.1
	improved code by dennis koepke

*)
END_FUNCTION

(* ---- CSET.st ---- *)
FUNCTION CSET : complex
VAR_INPUT
    RE : REAL;
    IM : REAL;
END_VAR
CSET.re := RE;
CSET.im := IM;

(* revision history
hm	21. feb 2008	rev 1.0
	original version

*)
END_FUNCTION

(* ---- CSIN.st ---- *)
FUNCTION CSIN : complex
VAR_INPUT
    X : complex;
END_VAR
CSIN.re := cosH(X.im) * SIN(X.re);
CSIN.im := sinH(X.im) * COS(X.re);

(* revision history
hm	21. feb 2008	rev 1.0
	original version

*)
END_FUNCTION

(* ---- CSINH.st ---- *)
FUNCTION CSINH : complex
VAR_INPUT
    X : COMPLEX;
END_VAR
CSINH.re := sinH(X.re) * COS(X.im);
CSINH.im := cosH(X.re) * SIN(X.im);

(* revision history
hm	21. feb 2008	rev 1.0
	original version

*)
END_FUNCTION

(* ---- CSQRT.st ---- *)
FUNCTION CSQRT : complex
VAR_INPUT
    X : complex;
END_VAR

VAR
    temp : REAL;
END_VAR
temp := HYPOT(x.re, x.im);
CSQRT.re :=  SQRT(0.5 * (temp + x.re));
CSQRT.im :=  sgn(x.im) * SQRT(0.5 * (temp - x.re));

(* revision history
hm	21. feb 2008	rev 1.0
	original version

*)
END_FUNCTION

(* ---- CSUB.st ---- *)
FUNCTION CSUB : complex
VAR_INPUT
    X : COMPLEX;
    Y : COMPLEX;
END_VAR
CSUB.re := X.re - Y.re;
CSUB.im := X.im - Y.im;

(* revision history
hm	21. feb 2008	rev 1.0
	original version

*)
END_FUNCTION

(* ---- CSV_PARSER_BUF_DEMO.st ---- *)
FUNCTION CSV_PARSER_BUF_DEMO
VAR_CONSTANT
    line_cnt : INT := 2;
    col_cnt : INT := 4;
END_VAR

VAR
    CPB : CSV_PARSER_BUF;
    FS : FILE_SERVER;
    FSD : FILE_SERVER_DATA;
    PT : NETWORK_BUFFER;
    sep : BYTE;
    value : STRING(OSCAT_BASIC.STRING_LENGTH);
    step : INT;
    result : BYTE;
    offset : UDINT;
    run : BYTE;
    done : BOOL;
    value_real : REAL;
    cnt : INT;
    line : INT;
    idx : INT;
    data : ARRAY[1..line_cnt, 1..col_cnt] OF REAL;
END_VAR
(* Demo-Programm: CSV-Datei mittels Enumeration auswerten
die groesse des arrays kann mittels konstanten line_cnt und col_cnt angepasst werden

 ----- den nachfolgenden Textblock als datei "csv.txt" auf der sps ablegen ---
10.45,20,30,40.8
115,3450.2123,456,123.1
---------------------------------------------------------------------------------*)

CASE step OF

00:	IF NOT done THEN
	 	(* File_Daten einrichten  *)
		FSD.FILENAME := 'csv.txt'; (* Dateiname *)
		FSD.MODE := 1; (* vorhandene Datei zum lesen öffnen *)
		FSD.OFFSET := 0; (* Start bei Dateianfang *)
		PT.SIZE := 65535; (* maximale länge einlesen *)
		step := 10;
	END_IF;

10:	IF FSD.MODE = 0 THEN (* Datei geöffnet ? *)
		OFFSET := 0; (* Start Offset vorgeben *)
		sep :=44; (* Trennzeichen , *)
		run := 1; (* Element suchen *)
		cnt := 0;
		step := 20;
	END_IF;

20:	IF run = 0 THEN
		(* ---------------------- Debug-Message ----------------------------*)
		(*IF _debug_enable THEN
			LOG_CL.NEW_MSG := 'CPFD: /value >~2< /offset ~3 /Run ~4 /Result ~5';
			LOG_CL.PRINTF[2] := value;
			LOG_CL.PRINTF[3] := UDINT_TO_STRING(OFFSET);
			LOG_CL.PRINTF[4] := BYTE_TO_STRING(run);
			LOG_CL.PRINTF[5] := BYTE_TO_STRING(result);
			LOG_MSG();
		END_IF;*)
		(* -----------------------------------------------------------------*)

		run := 1; (*  nächstes Element suchen  *)

		IF result = 1 OR result = 2 THEN
			(* automatische konvertierung in real ausführen *)
			IF LEN(value) <= 20 THEN
				value_real := OSCAT_BASIC.FLOAT_TO_REAL(FLT:=value);
			ELSE
				value_real := 0.0;
			END_IF;

			cnt := cnt + 1;
			IF cnt <= line_cnt * col_cnt THEN
				line := (cnt / col_cnt) + 1;
				idx := (cnt MOD col_cnt);
				data[line,idx] := value_real; (* Daten in Array eintragen *)
			END_IF;

		ELSIF result = 10 THEN (* nichts mehr gefunden *)
			run := 0; (* keine weitere INI Auswertung erwünscht *)
			FSD.MODE := 5; (* Datei schliessen *)
			step := 30;
		END_IF;
	END_IF;

30:	IF FSD.MODE = 0 THEN (* Datei geschlossen ? *)
		step := 0;
		done := TRUE;
	END_IF;

END_CASE;

CPB(SEP:=sep,RUN:=run,OFFSET:=OFFSET,VALUE:=value,PT:=PT,RESULT=>result); (* CSV PARAMETER BUF *)
FS(FSD:=FSD,PT:=PT); (* FILE_SERVER *)
END_FUNCTION

(* ---- CSV_PARSER_FILE_DEMO.st ---- *)
FUNCTION CSV_PARSER_FILE_DEMO
VAR CONSTANT
    line_cnt : INT := 2;
    col_cnt : INT := 4;
END_VAR

VAR
    CPF : CSV_PARSER_FILE;
    FS : FILE_SERVER;
    FSD : FILE_SERVER_DATA;
    PT : NETWORK_BUFFER;
    filename : STRING;
    value : STRING[OSCAT_BASIC.STRING_LENGTH];
    sep : BYTE;
    step : INT;
    result : BYTE;
    offset : UDINT;
    run : BYTE;
    done : BOOL;
    value_real : REAL;
    cnt : INT;
    line : INT;
    idx : INT;
    data : ARRAY[1..line_cnt, 1..col_cnt] OF REAL;
END_VAR
(* Demo-Programm: CSV-Datei mittels Enumeration auswerten

die groesse des arrays kann mittels konstanten line_cnt und col_cnt angepasst werden

 ----- den nachfolgenden Textblock als datei "csv.txt" auf der sps ablegen ---
10.45,20,30,40.8
115,3450.2123,456,123.1
---------------------------------------------------------------------------------*)

CASE step OF

00:	IF NOT done THEN
		filename := 'csv.txt'; (* File_Daten einrichten *)
		OFFSET := 0; (* Start Offset vorgeben *)
		sep :=44; (* Trennzeichen , *)
		run := 1; (* Element suchen *)
		cnt := 0;
		step := 20;
	END_IF;

20:	IF run = 0 THEN (* kein Befehl mehr aktiv ? *)
		(* ---------------------- Debug-Message ----------------------------*)
		(*IF _debug_enable THEN
			LOG_CL.NEW_MSG := 'CPFD: /value >~2< /offset ~3 /Run ~4 /Result ~5';
			LOG_CL.PRINTF[2] := value;
			LOG_CL.PRINTF[3] := UDINT_TO_STRING(OFFSET);
			LOG_CL.PRINTF[4] := BYTE_TO_STRING(run);
			LOG_CL.PRINTF[5] := BYTE_TO_STRING(result);
			LOG_MSG();
		END_IF;*)
		(* -----------------------------------------------------------------*)

		run := 1; (*  nächstes Element suchen  *)

		IF result = 1 OR result = 2 THEN
			(* automatische konvertierung in real ausführen *)
			IF LEN(value) <= 20 THEN
				value_real := OSCAT_BASIC.FLOAT_TO_REAL(FLT:=value);
			ELSE
				value_real := 0.0;
			END_IF;

			cnt := cnt + 1;
			IF cnt <= line_cnt * col_cnt THEN
				line := (cnt / col_cnt) + 1;
				idx := (cnt MOD col_cnt);
				data[line,idx] := value_real; (* Daten in Array eintragen *)
			END_IF;

		ELSIF result = 10 THEN (* nichts mehr gefunden *)
			run := 0; (* keine weitere INI Auswertung erwünscht *)
			FSD.MODE := 5; (* Datei schliessen *)
			step := 30;
		END_IF;
	END_IF;

30:	IF FSD.MODE = 0 THEN (* Befehl Datei schliessen beendet *)
		step := 0;
		done := TRUE;
	END_IF;

END_CASE;

CPF(SEP:=sep,FILENAME:=FILENAME,FSD:=FSD,RUN:=run,OFFSET:=OFFSET,VALUE:=value,PT:=PT,RESULT=>result); (* CSV PARAMETER FILE *)
FS(FSD:=FSD,PT:=PT); (* FILE_SERVER *)
END_FUNCTION

(* ---- CTAN.st ---- *)
FUNCTION CTAN : complex
VAR_INPUT
    X : complex;
END_VAR

VAR
    temp : REAL;
    xi2 : REAL;
    xr2 : REAL;
END_VAR
xi2 := 2.0 * x.im;
xr2 := 2.0 * x.re;
temp := 1.0 / (COS(xr2) + COSH( xi2));
CTAN.re := temp * SIN(xr2);
CTAN.im := temp * SINH(xi2);

(* revision history
hm	21. feb 2008	rev 1.0
	original version

hm	10. mar 2009	rev 1.1
	faster code
*)
END_FUNCTION

(* ---- CTANH.st ---- *)
FUNCTION CTANH : complex
VAR_INPUT
    X : complex;
END_VAR

VAR
    temp : REAL;
    xi2 : REAL;
    xr2 : REAL;
END_VAR
xi2 := 2.0 * x.im;
xr2 := 2.0 * x.re;
temp := 1.0 / (COSH(xr2) + COS(xi2));
CTANH.re := temp * SINH(xr2);
CTANH.im := temp * SIN(xi2);

(* revision history
hm	21. feb 2008	rev 1.0
	original version

hm	10. mar. 2009	rev 1.1
	new faster code

*)
END_FUNCTION

(* ---- CTRL_IN.st ---- *)
FUNCTION CTRL_IN : REAL
VAR_INPUT
    SET_POINT : REAL;
    ACTUAL : REAL;
    NOISE : REAL;
END_VAR
(* calculate the process error DIFF *)
CTRL_IN := DEAD_ZONE(SET_POINT - ACTUAL, NOISE);

(* revision history
hm 	2. jun. 2008 	rev 1.0
	original version

*)
END_FUNCTION

(* ---- D_TRUNC.st ---- *)
FUNCTION D_TRUNC : DINT
VAR_INPUT
    X : REAL;
END_VAR
D_TRUNC := REAL_TO_DINT(X);
IF X > 0.0 THEN
	IF DINT_TO_REAL(D_TRUNC) > X THEN D_TRUNC := D_TRUNC - 1; END_IF;
ELSE
	IF DINT_TO_REAL(D_TRUNC) < X THEN D_TRUNC := D_TRUNC + 1; END_IF;
END_IF;

(* for systems that support a dint truncation this routine can be replaced by trunc() *)

(* revision history
hm	21. mar. 2008	rev 1.0
	original version

hm	31. oct. 2008	rev 1.1
	optimized performance

hm	10. mar. 2009	rev 1.2
	real constants updated to new systax using dot
*)
END_FUNCTION

(* ---- DATE_ADD.st ---- *)
FUNCTION DATE_ADD : DATE
VAR_INPUT
    IDATE: DATE;
    D: INT;
    W: INT;
    M: INT;
    Y: INT;
END_VAR

VAR
    mo: INT;
    yr: INT;
    dm: INT;
END_VAR
DATE_ADD := UDINT_TO_DATE(DATE_TO_UDINT(IDATE) + INT_TO_UDINT(D + W * 7) * UDINT#86400);
yr := Y + YEAR_OF_DATE(DATE_ADD);
mo := M + MONTH_OF_DATE(DATE_ADD);
dm := DAY_OF_MONTH(DATE_ADD);
WHILE mo > 12 DO
	mo := mo - 12;
	yr := yr + 1;
END_WHILE;
WHILE mo < 1 DO
	mo := mo + 12;
	yr := yr - 1;
END_WHILE;
DATE_ADD := SET_DATE(yr, mo, dm);

(* revision history

hm 27.12.2006	rev 1.0
	nrw module

hm 12.4.2007		rev 1.1
	corrected an error while date would be incorrect when year  = 0

hm	1.11.2007		rev 1.2
	added int_to_dword stetements to avoid possible overrun with möller ecp4

hm	22. mar. 2008	rev 1.3
	fixed some bugs when month was negative

hm	7. oct. 2008	rev 1.4
	changed function year to year_of_date
	changed function month to month_of_date

hm	29. mar. 2009	rev 1.5
	improved performance

hm	27. jan. 2011	rev 1.6
	faster code

hm	2. feb. 2011		rev 1.7
	fixed an error, weeks not calculated

hm	22. mar. 2011	rev 1.8
	fixed an error in formula
*)
END_FUNCTION

(* ---- DAY_OF_DATE.st ---- *)
FUNCTION DAY_OF_DATE : DINT
VAR_INPUT
    idate : DATE;
END_VAR
DAY_OF_DATE := DWORD_TO_DINT(DATE_TO_DWORD(idate) / 86400);

(* revision history
hm		16.9.2007		rev 1.0
	original version

hm		1. okt 2007		rev 1.1
	added step7 compatibility

hm		22. mar. 2008	rev 1.2
	changed output from int to Dint because the total date range is 49710 days

hm		7. apr. 2008	rev 1.3
	deleted unused step7 code

*)
END_FUNCTION

(* ---- DAY_OF_MONTH.st ---- *)
FUNCTION DAY_OF_MONTH : INT
VAR_INPUT
    IDATE : DATE;
END_VAR

VAR
    leap : INT;
END_VAR
(* calculate the day in the year *)
DAY_OF_MONTH := DAY_OF_YEAR(idate);
(* leap will be set to one for a leap year *)
leap := BOOL_TO_INT(LEAP_OF_DATE(idate));
(* if leap year deduct one from the days of the year *)
DAY_OF_MONTH := DAY_OF_MONTH - leap;
(* search if we are in month december to march ? *)
IF DAY_OF_MONTH > setup.MTH_OFS[9] THEN
	IF DAY_OF_MONTH > setup.MTH_OFS[11] THEN
		IF DAY_OF_MONTH > setup.mth_ofs[12] THEN
			DAY_OF_MONTH := DAY_OF_MONTH - setup.MTH_OFS[12];
		ELSE
			DAY_OF_MONTH := DAY_OF_MONTH - setup.MTH_OFS[11];
		END_IF;
	ELSE
		IF DAY_OF_MONTH > setup.mth_ofs[10] THEN
			DAY_OF_MONTH := DAY_OF_MONTH - setup.MTH_OFS[10];
		ELSE
			DAY_OF_MONTH := DAY_OF_MONTH - setup.MTH_OFS[9];
		END_IF;
	END_IF;
ELSIF DAY_OF_MONTH > setup.MTH_OFS[5] THEN
	IF DAY_OF_MONTH > setup.MTH_OFS[7] THEN
		IF DAY_OF_MONTH > setup.mth_ofs[8] THEN
			DAY_OF_MONTH := DAY_OF_MONTH - setup.MTH_OFS[8];
		ELSE
			DAY_OF_MONTH := DAY_OF_MONTH - setup.MTH_OFS[7];
		END_IF;
	ELSE
		IF DAY_OF_MONTH > setup.mth_ofs[6] THEN
			DAY_OF_MONTH := DAY_OF_MONTH - setup.MTH_OFS[6];
		ELSE
			DAY_OF_MONTH := DAY_OF_MONTH - setup.MTH_OFS[5];
		END_IF;
	END_IF;
ELSIF DAY_OF_MONTH > setup.MTH_OFS[3] THEN
	IF DAY_OF_MONTH > setup.MTH_OFS[4] THEN
		DAY_OF_MONTH := DAY_OF_MONTH - setup.MTH_OFS[4];
	ELSE
		DAY_OF_MONTH := DAY_OF_MONTH - setup.MTH_OFS[3];
	END_IF;
ELSE
	(* since now we must be in february or january we need to add leap again *)
	DAY_OF_MONTH := DAY_OF_MONTH + leap;
	IF DAY_OF_MONTH > setup.MTH_OFS[2] THEN DAY_OF_MONTH := DAY_OF_MONTH - setup.mth_ofs[2]; END_IF;
	(* since nothing was true before, day_of_month must already be good *)
END_IF;

(*
Revision history

hm 22.1.2007		rev 1.1
	deleted unused variable day_in_year and day_in_year_begin

hm	1. okt 2007	rev 1.2
	changed code to use day_of_year and leap_of_date
	added compatibility to STEP7

hm	8. oct 2007	rev 1.3
	deleted unused variable yr

hm	8. jan 2008	rev 1.4
	improved performance

hm	25. oct. 2008	rev 2.0
	new code using setup constants

hm	10. mar. 2009	rev 2.1
	removed nested comments

*)
END_FUNCTION

(* ---- DAY_OF_WEEK.st ---- *)
FUNCTION DAY_OF_WEEK : INT
VAR_INPUT
    IDATE: DATE;
END_VAR
DAY_OF_WEEK := DWORD_TO_INT((DATE_TO_DWORD(idate) / 86400 + 3) MOD 7) + 1;

(* revision history
hm 	21.8.06 		rev 1.1
	corrected a miscalculation

hm	23.12.2007		rev 1.2
	correction for step7

hm	7. apr. 2008	rev 1.3
	deleted unused step7 code

hm	7. oct. 2008	rev 1.4
	changed name of function from weekday to day_of_week

*)
END_FUNCTION

(* ---- DAY_OF_YEAR.st ---- *)
FUNCTION DAY_OF_YEAR : INT
VAR_INPUT
    IDATE : DATE;
END_VAR
DAY_OF_YEAR := UDINT_TO_INT((DATE_TO_UDINT(idate) / UDINT#86400) MOD UDINT#1461);
IF DAY_OF_YEAR > 729 THEN
	IF DAY_OF_YEAR > 1095 THEN DAY_OF_YEAR := DAY_OF_YEAR - 1095; ELSE DAY_OF_YEAR := DAY_OF_YEAR - 729; END_IF;
ELSIF DAY_OF_YEAR > 364 THEN
	DAY_OF_YEAR := DAY_OF_YEAR - 364;
ELSE
	DAY_OF_YEAR := DAY_OF_YEAR + 1;
END_IF;

(*
DAY_OF_YEAR := DWORD_TO_INT((DATE_TO_DWORD(idate) - DATE_TO_DWORD(YEAR_BEGIN(YEAR_OF_DATE(idate)))) / 86400) + 1;
*)

(* revivision history
hm	4. aug. 2007		rev 1.0
	original version

hm	1. oct. 2007		rev 1.1
	added compatibility to STEP7

hm	4. jan. 2008		rev 1.2
	changed code for better performance

hm	7. oct. 2008		rev 1.3
	changed name of function year to year_of_date

hm	28. jan. 2011	rev 1.4
	improved code
*)
END_FUNCTION

(* ---- DAY_TO_TIME.st ---- *)
FUNCTION DAY_TO_TIME : TIME
VAR_INPUT
    IN : REAL;
END_VAR
DAY_TO_TIME := DWORD_TO_TIME(REAL_TO_DWORD(IN * 86400000.0));

(* revision history
hm	4. aug. 2006	rev 1.0
	original release

hm	24. feb. 2009	rev 1.1
	renamed input to IN
*)
END_FUNCTION

(* ---- DAYS_DELTA.st ---- *)
FUNCTION DAYS_DELTA : DINT
VAR_INPUT
    date_1 : DATE;
    date_2 : DATE;
END_VAR
IF DATE_1 > DATE_2 THEN
	DAYS_DELTA := - DWORD_TO_DINT((DATE_TO_DWORD(date_1) - DATE_TO_DWORD(date_2)) / 86400);
ELSE
	DAYS_DELTA := DWORD_TO_DINT((DATE_TO_DWORD(date_2) - DATE_TO_DWORD(date_1)) / 86400);
END_IF;

(* revision history
hm	27. dec 2006	rev 1.0
	original version

hm	16.9.2007		rev 1.1
	coorected an error in formula and changed algorithm to show positive and negative delta

hm	22. mar. 2008	rev 1.2
	changed output from int to dint because the total date range is 49710 days

hm	25. jan. 2011	rev 1.3
	improved performance
*)
END_FUNCTION

(* ---- DAYS_IN_MONTH.st ---- *)
FUNCTION DAYS_IN_MONTH : INT
VAR_INPUT
    IDATE : DATE;
END_VAR
DAYS_IN_MONTH := DAY_OF_YEAR(IDATE);
IF LEAP_OF_DATE(IDATE) THEN
	CASE DAYS_IN_MONTH OF
		32..60	:	DAYS_IN_MONTH := 29;
		92..121 :	DAYS_IN_MONTH := 30;
		153..182:	DAYS_IN_MONTH := 30;
		245..274:	DAYS_IN_MONTH := 30;
		306..335:	DAYS_IN_MONTH := 30;
	ELSE
		DAYS_IN_MONTH := 31;
	END_CASE;
ELSE
	CASE DAYS_IN_MONTH OF
		32..59	:	DAYS_IN_MONTH := 28;
		91..120 :	DAYS_IN_MONTH := 30;
		152..181:	DAYS_IN_MONTH := 30;
		244..273:	DAYS_IN_MONTH := 30;
		305..334:	DAYS_IN_MONTH := 30;
	ELSE
		DAYS_IN_MONTH := 31;
	END_CASE;
END_IF;

(* revision history
hm	27. mar. 2009		rev 1.0
	original version

*)
END_FUNCTION

(* ---- DAYS_IN_YEAR.st ---- *)
FUNCTION DAYS_IN_YEAR : INT
VAR_INPUT
    IDATE : DATE;
END_VAR
IF LEAP_OF_DATE(IDATE) THEN
	DAYS_IN_YEAR := 366;
ELSE
	DAYS_IN_YEAR := 365;
END_IF;

(* revision history
hm	27. mar. 2009		rev 1.0
	original version

*)
END_FUNCTION

(* ---- DEAD_BAND.st ---- *)
FUNCTION DEAD_BAND : REAL
VAR_INPUT
    X : REAL;
    L : REAL;
END_VAR
IF X > L THEN
	DEAD_BAND := X - L;
ELSIF X < -L THEN
	DEAD_BAND := X + L;
ELSE
	DEAD_BAND := 0.0;
END_IF;

(* revision history
hm	2. nov. 2007	rev 1.0
	original version

hm	14. jun. 2008	rev 1.1
	improved performance

hm	18. jan. 2011	rev 1.2
	assign 0 before return
*)
END_FUNCTION

(* ---- DEAD_ZONE.st ---- *)
FUNCTION DEAD_ZONE : REAL
VAR_INPUT
    X : REAL;  // Input variable X of type REAL
    L : REAL;  // Input variable L of type REAL
END_VAR
IF ABS(x) > L THEN
	dead_zone := X;
ELSE
	DEAD_ZONE := 0.0;
END_IF;

(* revision history
hm	12. feb. 2007	rev 1.0
	original version

hm	14. jun. 2008	rev 1.1
	improved performance

hm	11. mar. 2009	rev 1.2
	real constants updated to new systax using dot

*)
END_FUNCTION

(* ---- DEC1.st ---- *)
FUNCTION DEC1 : INT
VAR_INPUT
    X : INT;
    N : INT;
END_VAR
IF X = 0 THEN
	DEC1 := N - 1;
ELSE
	DEC1 := X - 1;
END_IF;

(* this is a very elegant version but 50% slower
X := (X - 1 + N) MOD N;
*)

(* revision history
hm	13. oct. 2008	rev 1.0
	original version

hm	27. oct. 2008	rev 1.1
	added statement to return value for compatibility reasons

*)
END_FUNCTION

(* ---- DEC_TO_BYTE.st ---- *)
FUNCTION DEC_TO_BYTE : BYTE
VAR_INPUT
    DEC : STRING(10);
END_VAR

VAR
    pt : POINTER TO BYTE;
    i : INT;
    X : BYTE;
    stop : INT;
END_VAR
pt := ADR(dec);
stop := LEN(DEC);
FOR I := 1 TO stop DO
	(* read the first character and subtract 48 to get value in decimal 0 = 48 *)
	x := pt^;
	(* calculate the value of the digit *)
	IF X > 47 AND x < 58 THEN
		DEC_TO_BYTE := DEC_TO_BYTE * 10 + X - 48;
	END_IF;
	pt := pt + 1;
END_FOR;

(* revision histroy
hm	20. jun. 2008	rev 1.0
	original release

hm	30. sep.2008	rev 1.1
	changed length of input string from 20 to 10
	corrected an error where decoding of characters 8 and 9 would fail

*)
END_FUNCTION

(* ---- DEC_TO_DWORD.st ---- *)
FUNCTION DEC_TO_DWORD : DWORD
VAR_INPUT
    DEC : STRING[20];
END_VAR

VAR
    pt : POINTER TO BYTE;
    i : INT;
    X : BYTE;
    stop : INT;
END_VAR
pt := ADR(dec);
stop := LEN(dec);
FOR I := 1 TO stop DO
	(* read the first character and subtract 48 to get value in decimal 0 = 48 *)
	x := pt^;
	(* calculate the value of the digit *)
	IF X > 47 AND x < 58 THEN
		DEC_TO_DWORD := DEC_TO_DWORD * 10 + X - 48;
	END_IF;
	pt := pt + 1;
END_FOR;

(* revision histroy
hm	20. jun. 2008	rev 1.0
	original release

hm	30. sep. 2008	rev 1.1
	corrected an error where decoding of characters 8 and 9 would fail
*)
END_FUNCTION

(* ---- DEC_TO_INT.st ---- *)
FUNCTION DEC_TO_INT : INT
VAR_INPUT
    DEC: STRING[10];
END_VAR

VAR
    pt: POINTER TO BYTE;
    i: INT;
    X: BYTE;
    sign: BOOL;
    stop: INT;
END_VAR
pt := ADR(dec);
stop := LEN(dec);
FOR I := 1 TO stop DO
	(* read the first character and subtract 48 to get value in decimal 0 = 48 *)
	x := pt^;
	(* calculate the value of the digit *)
	IF X > 47 AND x < 58 THEN
		DEC_TO_INT := DEC_TO_INT * 10 + X - 48;
	ELSIF X = 45 AND DEC_TO_INT = 0 THEN
		sign := TRUE;
	END_IF;
	pt := pt + 1;
END_FOR;
IF sign THEN DEC_TO_INT := -DEC_TO_INT; END_IF;

(* revision histroy
hm	20. jun. 2008	rev 1.0
	original release

hm	30. sep. 2008	rev 1.1
	changed length of input string from 20 to 10
	corrected an error where decoding of characters 8 and 9 would fail
*)
END_FUNCTION

(* ---- DEG.st ---- *)
FUNCTION DEG : REAL
VAR_INPUT
    rad : REAL;
END_VAR
DEG := MODR(57.29577951308232 * RAD, 360.0);

(* revision history
hm	4. aug 2006	rev 1.0
	original version

hm 16. oct 2007	rev 1.1
	added modr statement which prohibits deg to become bigger than 360

hm	10. mar. 2009	rev 1.2
	real constants updated to new systax using dot
*)
END_FUNCTION

(* ---- DEG_TO_DIR.st ---- *)
FUNCTION DEG_TO_DIR : string
VAR_INPUT
    DEG : INT;  // Degree input
    N   : INT;  // Another input variable
    L   : INT;  // Length input
END_VAR

VAR
    ly  : INT;  // Local variable
END_VAR
IF L = 0 THEN ly := LANGUAGE.DEFAULT; ELSE ly := MIN(L, LANGUAGE.LMAX); END_IF;
DEG_TO_DIR := LANGUAGE.DIRS[ly, ((SHL(DEG,N-1) + 45) / 90) MOD SHL(INT#2,N)*SHR(INT#8,N)];

(*
DIR := ((SHL(DEG,N-1) + 45) / 90) MOD SHL(INT#2,N);
explanation :
DIR is calculated BY the following formula:
DIR := ((DIR + 45) / 90) MOD 4 if N = 1 digit
North = 0, East = 1 ....
DIR := ((DIR + 22,5) / 45) MOD 8 if N = 2 digit
convert to integer calculation
DIR := ((DIR*2 + 45) / 90) MOD 8
N = 0, NE = 1 ....
ther above formula replaces 2^N with shift for performance
*)

(* revision histroy
hm	11. jun. 2008	rev 1.0
	original release

hm	22. oct. 2008	rev 1.1
	changed size of string variables to 30
*)
END_FUNCTION

(* ---- DEL_CHARS.st ---- *)
FUNCTION DEL_CHARS : string
VAR_INPUT
    IN : STRING; // Length not specified in ST code
    CX : STRING[80];
END_VAR

VAR
    pos : INT := 1;
    stop : INT;
END_VAR
(* copy input string *)
DEL_CHARS := IN;
stop := LEN(in);
WHILE pos <= stop DO
	IF FIND(cx, MID(DEL_CHARS, 1, pos)) > 0 THEN
		(* wrong chracter needs to be deleted *)
		DEL_CHARS := DELETE(DEL_CHARS, 1, pos);
		stop := stop - 1;	(* the string is one character shorter now *)
	ELSE
		(* charcter not found skip to next one *)
		pos := pos + 1;
	END_IF;
END_WHILE;

(* revision history

hm		18. jun. 2008	rev 1.0
	original version

*)
END_FUNCTION

(* ---- DEW_CON.st ---- *)
FUNCTION DEW_CON : REAL
VAR_INPUT
    RH : REAL; // Relative Humidity
    T : REAL;  // Temperature
END_VAR
(*	this code is good to read but need to be improoved
	SDD := 6.1078*EXPT(10,(a*T)/(b+T));
	DD := RH/100 * SDD;
	V := LOG(DD/6.1078);
	TD := b*V/(a-v);
	dew_con := 0.1 * mw / RU * DD / (T - TK);
*)
IF RH > 0.0 AND T > -50.0 THEN
	DEW_CON := 2.166824303E-2 * RH * SDD(T,FALSE)  / (T - OSCAT_BASIC.phys.T0);
ELSE
	DEW_CON := 0.0;
END_IF;

(*
Bezeichnungen:
r = relative Luftfeuchte
T = Temperatur in °C
TK = Temperatur in Kelvin (TK = T + 273.15)
TD = Taupunkttemperatur in °C
DD = Dampfdruck in hPa
SDD = Sättigungsdampfdruck in hPa

Parameter:
a = 7.5, b = 237.3 für T >= 0
a = 7.6, b = 240.7 für T < 0 über Wasser (Taupunkt)
a = 9.5, b = 265.5 für T < 0 über Eis (Frostpunkt)

R* = 8314.3 J/(kmol*K) (universelle Gaskonstante)
mw = 18.016 kg (Molekulargewicht des Wasserdampfes)
AF = absolute Feuchte in g Wasserdampf pro m3 Luft

Formeln:

   1. SDD(T) = 6.1078 * 10^((a*T)/(b+T))
   2. DD(r,T) = r/100 * SDD(T)
   3. r(T,TD) = 100 * SDD(TD) / SDD(T)
   4. TD(r,T) = b*v/(a-v) mit v(r,T) = log10(DD(r,T)/6.1078)
   5. AF(r,TK) = 10^5 * mw/R* * DD(r,T)/TK; AF(TD,TK) = 10^5 * mw/R* * SDD(TD)/TK

*)

(* revision history

hm 29 apr 2007	rev 1.0
	original version

hm	13.sep 2007	rev 1.1
	improoved coding for speed
	deleted unused variabled SDD,DD,V, TD

hm	2. dec 2007	rev 1.2
	changed code for better performance
	output is now in Gramms / Qubic meter

hm	14. oct. 2008	rev 1.3
	performance improvement

hm	18. oct. 2008	rev 1.4
	using phys constants

hm	13. mar. 2009	rev 1.5
	improved code

hm	19. jan. 2011	rev 1.6
	return value 0.0 if RH <= 0.0

*)
END_FUNCTION

(* ---- DEW_RH.st ---- *)
FUNCTION DEW_RH : REAL
VAR_INPUT
    VC : REAL;
    T : REAL;
END_VAR
DEW_RH := LIMIT(0.0, VC / DEW_CON(1.0, T), 100.0);

(* code before rev 1.1
dew_rh := VC / dew_con(100,T) * 100;
IF dew_rh > 100 THEN dew_rh := 100; END_IF;
*)

(* revision history
hm	29. apr 2007	rev 1.0
	original version

hm	2. 12. 2007	rev 1.1
	new code for better performance

hm	13. mar. 2009	rev 1.2
	real constants updated to new systax using dot

*)
END_FUNCTION

(* ---- DEW_TEMP.st ---- *)
FUNCTION DEW_TEMP : REAL
VAR_INPUT
    RH : REAL;
    T : REAL;
END_VAR

VAR CONSTANT
    a : REAL := 7.5;
    b : REAL := 237.3;
END_VAR

VAR
    V : REAL;
END_VAR
IF rh > 0.0 THEN
(*	old code was rewritten for better performance
	SDD := 6.1078*EXPT(10,(a*T)/(b+T));
	DD := RH/100 * SDD;
	V := LOG(DD/6.1078);
	dew_temp := b*V/(a-v);
*)
	V := LOG(RH * 0.01 * OSCAT_BASIC.EXP10((a*T) / (b+T)));
	DEW_TEMP := b*V / (a-V);
ELSE
	DEW_TEMP:= OSCAT_BASIC.phys.T0;
END_IF;

(* revision history

hm		2.10.2006	rev 1.0
	original version created

hm		29.4.2007	rev 1.1
	checked for rh not to be 0 because log(0) is not defined

hm		13.9.2007	rev 1.2
	code rewritten for better performance

hm	2. dec 2007	rev 1.3
	changed code for better performance

hm	8. jan 2008	rev 1.4
	further improvement in performance

hm	18. oct. 2008	rev 1.5
	using phys constants

hm	13. mar. 2009	rev 1.6
	real constants updated to new systax using dot
	function will now return -273.15 °C for RH = 0
*)

(*
Bezeichnungen:
r = relative Luftfeuchte
T = Temperatur in °C
TK = Temperatur in Kelvin (TK = T + 273.15)
TD = Taupunkttemperatur in °C
DD = Dampfdruck in hPa
SDD = Sättigungsdampfdruck in hPa

Parameter:
a = 7.5, b = 237.3 für T >= 0
a = 7.6, b = 240.7 für T < 0 über Wasser (Taupunkt)
a = 9.5, b = 265.5 für T < 0 über Eis (Frostpunkt)

R* = 8314.3 J/(kmol*K) (universelle Gaskonstante)
mw = 18.016 kg (Molekulargewicht des Wasserdampfes)
AF = absolute Feuchte in g Wasserdampf pro m3 Luft

Formeln:

   1. SDD(T) = 6.1078 * 10^((a*T)/(b+T))
   2. DD(r,T) = r/100 * SDD(T)
   3. r(T,TD) = 100 * SDD(TD) / SDD(T)
   4. TD(r,T) = b*v/(a-v) mit v(r,T) = log10(DD(r,T)/6.1078)
   5. AF(r,TK) = 10^5 * mw/R* * DD(r,T)/TK; AF(TD,TK) = 10^5 * mw/R* * SDD(TD)/TK

*)
END_FUNCTION

(* ---- DIFFER.st ---- *)
FUNCTION DIFFER : BOOL
VAR_INPUT
    in1 : REAL;
    in2 : REAL;
    X : REAL;
END_VAR
DIFFER := ABS(in1 - in2) > X;

(* revision history
hm		8. oct 2006		rev 1.0
	original version

hm		16. mar 2008	rev 1.1
	improverd code for performance

*)
END_FUNCTION

(* ---- DIR_TO_DEG.st ---- *)
FUNCTION DIR_TO_DEG : INT
VAR_INPUT
    DIR: STRING[3];
    L: INT;
END_VAR

VAR
    ly: INT;
    i: INT;
END_VAR
IF L = 0 THEN ly := LANGUAGE.DEFAULT; ELSE ly := MIN(L, LANGUAGE.LMAX); END_IF;
FOR i := 0 TO 15 DO
	IF language.DIRS[ly, i] = DIR THEN EXIT; END_IF;
END_FOR;
DIR_TO_DEG := SHR(i * 45 + 1, 1);

(* revision histroy
hm	22. oct. 2008	rev 1.1
	original release

*)
END_FUNCTION

(* ---- DLOG_FILE_CSV_DEMO.st ---- *)
FUNCTION DLOG_FILE_CSV_DEMO
VAR
    cur_dt: DT;
    enable: BOOL := TRUE;
    trig_t: TIME := TIME#5s0ms;
    trig_m: BOOL;
    error_c: DWORD;
    error_t: BYTE;
    auto_close: TIME := TIME#10s0ms;
    x1: DLOG_DT;
    x2: DLOG_REAL;
    x3: DLOG_DINT;
    x4: DLOG_BOOL;
    x5: DLOG_STRING;
    x: DLOG_DATA;
    RTC_2: oscat_basic.RTC_2;
    DLOG_STORE_FILE_CSV: DLOG_STORE_FILE_CSV;
    GEN_SIN_1: oscat_basic.GEN_SIN;
    COUNT_DR: oscat_basic.COUNT_DR;
    save_data: DLOG_SAVE; (* Retain variable *)
END_VAR

END_FUNCTION

(* ---- DLOG_FILE_CSV_FTP_DEMO.st ---- *)
FUNCTION DLOG_FILE_CSV_FTP_DEMO
VAR
    cur_dt: DT;
    enable: BOOL := TRUE;
    trig_t: TIME := TIME#5s0ms;
    trig_m: BOOL;
    error_c: DWORD;
    error_t: BYTE;
    auto_close: TIME := TIME#10s0ms;
    x1: DLOG_DT;
    x2: DLOG_REAL;
    x3: DLOG_DINT;
    x4: DLOG_BOOL;
    x5: DLOG_STRING;
    x: DLOG_DATA;
    RTC_2: oscat_basic.RTC_2;
    DLOG_STORE_FILE_CSV: DLOG_STORE_FILE_CSV;
    GEN_SIN_1: oscat_basic.GEN_SIN;
    COUNT_DR: oscat_basic.COUNT_DR;
    DLOG_FILE_TO_FTP: DLOG_FILE_TO_FTP;
    ftp_done: BOOL;
    ftp_busy: BOOL;
    ftp_error_c: DWORD;
    ftp_error_t: BYTE;
    ftp_url: STRING := 'ftp://581920:123456@oscat.atwebpages.com:2000/subordner/';
    ftp_activ: BOOL := FALSE;
    ftp_delete: BOOL := TRUE;
    ftp_retry: INT := 0;
    ftp_retry_time: TIME := TIME#1m0s0ms;
    ftp_timeout: TIME := TIME#30s0ms;
    save_data: DLOG_SAVE; // Retained variable
END_VAR

END_FUNCTION

(* ---- DLOG_FILE_CSV_SMTP_DEMO.st ---- *)
FUNCTION DLOG_FILE_CSV_SMTP_DEMO
VAR
    cur_dt : DT;
    enable : BOOL := TRUE;
    trig_t : TIME := TIME#5s0ms;
    trig_m : BOOL;
    error_c : DWORD;
    error_t : BYTE;
    auto_close : TIME := TIME#10s0ms;
    x1 : DLOG_DT;
    x2 : DLOG_REAL;
    x3 : DLOG_DINT;
    x4 : DLOG_BOOL;
    x5 : DLOG_STRING;
    x : DLOG_DATA;
    RTC_2 : oscat_basic.RTC_2;
    DLOG_STORE_FILE_CSV : DLOG_STORE_FILE_CSV;
    GEN_SIN_1 : oscat_basic.GEN_SIN;
    COUNT_DR : oscat_basic.COUNT_DR;
    DLOG_FILE_TO_SMTP : DLOG_FILE_TO_SMTP;
    smtp_timeout : TIME := TIME#30s0ms;
    smtp_error_t : BYTE;
    smtp_error_c : DWORD;
    smtp_busy : BOOL;
    smtp_done : BOOL;
    smtp_dti : DT;
    smtp_dti_offset : INT := 60;
    smtp_server : STRING := '110876022:oscat123456@mail.gmx.net';
    smtp_mailfrom : STRING := 'oscat@gmx.net;Station_01';
    smtp_mailto : STRING[OSCAT_BASIC.STRING_LENGTH] := 'oscat@gmx.net';
    smtp_subject : STRING := 'Das ist der Betreff';
    smtp_body : STRING[OSCAT_BASIC.STRING_LENGTH] := 'Das ist der Email-Text';
    smtp_delete : BOOL := TRUE;
    smtp_retry : INT := 0;
    smtp_retry_time : TIME := TIME#1m0s0ms;
    save_data : DLOG_SAVE;
END_VAR

END_FUNCTION

(* ---- DLOG_FILE_HTML_DEMO.st ---- *)
FUNCTION DLOG_FILE_HTML_DEMO
VAR
    cur_dt : DT;
    enable : BOOL := TRUE;
    trig_t : TIME := TIME#5s0ms;
    trig_m : BOOL;
    error_c : DWORD;
    error_t : BYTE;
    auto_close : TIME := TIME#10s0ms;
    x1 : DLOG_DT;
    x2 : DLOG_REAL;
    x3 : DLOG_DINT;
    x4 : DLOG_BOOL;
    x5 : DLOG_STRING;
    x : DLOG_DATA;
    RTC_2 : oscat_basic.RTC_2;
    DLOG_STORE_FILE_HTML : DLOG_STORE_FILE_HTML;
    GEN_SIN_1 : oscat_basic.GEN_SIN;
    COUNT_DR : oscat_basic.COUNT_DR;
    html_caption : STRING := 'Das ist der Titel';
    html_tr_even : STRING := 'BGCOLOR=#B3B7FF';
    html_tr_odd : STRING := 'BGCOLOR=#E0E0E0';
    html_tr_head : STRING := 'BGCOLOR=#FFFF40';
    html_table : STRING := 'BORDER="1"';
END_VAR

VAR RETAIN
    save_data : DLOG_SAVE;
END_VAR

END_FUNCTION

(* ---- DLOG_FILE_XML_DEMO.st ---- *)
FUNCTION DLOG_FILE_XML_DEMO
VAR
    cur_dt: DT;
    enable: BOOL := TRUE;
    trig_t: TIME := TIME#5s0ms;
    trig_m: BOOL;
    error_c: DWORD;
    error_t: BYTE;
    auto_close: TIME := TIME#10s0ms;
    x1: DLOG_DT;
    x2: DLOG_REAL;
    x3: DLOG_DINT;
    x4: DLOG_BOOL;
    x5: DLOG_STRING;
    x: DLOG_DATA;
    RTC_2: oscat_basic.RTC_2;
    DLOG_STORE_FILE_XML: DLOG_STORE_FILE_XML;
    GEN_SIN_1: oscat_basic.GEN_SIN;
    COUNT_DR: oscat_basic.COUNT_DR;
    save_data: DLOG_SAVE; // Retain variable
END_VAR

END_FUNCTION

(* ---- DLOG_MYSQL_DEMO.st ---- *)
FUNCTION DLOG_MYSQL_DEMO
VAR
    cur_dt : DT;
    enable : BOOL := TRUE;
    trig_t : TIME := TIME#5s0ms;
    trig_m : BOOL;
    error_c : DWORD;
    error_t : BYTE;
    x1 : DLOG_DT;
    x2 : DLOG_REAL;
    x3 : DLOG_DINT;
    x4 : DLOG_BOOL;
    x5 : DLOG_STRING;
    x : DLOG_DATA;
    mysql_info : MYSQL_INFO;
    RTC_2 : oscat_basic.RTC_2;
    GEN_SIN_1 : oscat_basic.GEN_SIN;
    COUNT_DR : oscat_basic.COUNT_DR;
    DLOG_STORE_MYSQL : DLOG_STORE_MYSQL;
    url : STRING[OSCAT_BASIC.STRING_LENGTH] := 'myuser:mypassword@192.168.178.21';
    db_name : STRING[64] := 'oscat_db';
    tb_name : STRING[64] := 'oscat_tb';
    auto_delete : UDINT := 0;
    timeout : TIME := TIME#10s0ms;
END_VAR

END_FUNCTION

(* ---- DLOG_RRD_DEMO.st ---- *)
FUNCTION DLOG_RRD_DEMO
VAR
    cur_dt : DT;
    trig_t : TIME := TIME#50s0ms;
    trig_m : BOOL;
    rrd_error_c : DWORD;
    rrd_error_t : BYTE;
    rrd_enable : BOOL := TRUE;
    rrd_url : STRING(OSCAT_BASIC.STRING_LENGTH) := '192.168.178.21/rrd/test_rrd2.php?rrd_db=test.rrd&value=';
    rrd_timeout : TIME := TIME#5s0ms;
    RTC_2 : oscat_basic.RTC_2;
    DLOG_STORE_RRD : DLOG_STORE_RRD;
    x : DLOG_DATA;
    x1 : DLOG_DINT;
    x2 : DLOG_DINT;
    x3 : DLOG_REAL;
    x4 : DLOG_REAL;
    x5 : DLOG_REAL;
    x6 : DLOG_REAL;
    x7 : DLOG_REAL;
    GEN_SIN_1 : oscat_basic.GEN_SIN;
    GEN_SIN_2 : oscat_basic.GEN_SIN;
    GEN_SIN_3 : oscat_basic.GEN_SIN;
    GEN_RMP_1 : oscat_basic.GEN_RMP;
    GEN_RMP_2 : oscat_basic.GEN_RMP;
END_VAR

END_FUNCTION

(* ---- DNS_DYN_DEMO.st ---- *)
FUNCTION DNS_DYN_DEMO
VAR
    DNS_DYN : DNS_DYN;
    IP_C : IP_C;
    S_BUF : NETWORK_BUFFER;
    R_BUF : NETWORK_BUFFER;
    IP_CONTROL : IP_CONTROL;
    enable : BOOL;
    done : BOOL;
    error_c : DWORD;
    error_t : BYTE;
    busy : BOOL;
    COUNT_DR : oscab_basic.COUNT_DR;
    z : DWORD;
    GET_WAN_IP : GET_WAN_IP;
    t1 : TON;
    done2 : BOOL;
    error_c2 : DWORD;
    error_t2 : BYTE;
    update : BOOL;
    new_ip : BOOL;
    wan_ip4 : DWORD;
END_VAR

END_FUNCTION

(* ---- DNS_REV_DEMO.st ---- *)
FUNCTION DNS_REV_DEMO
VAR
    DNS_REV_CLIENT : DNS_REV_CLIENT;
    IP_C : IP_C;
    S_BUF : NETWORK_BUFFER;
    R_BUF : NETWORK_BUFFER;
    IP_CONTROL : IP_CONTROL;
    activate : BOOL := TRUE;
    done : BOOL;
    error : DWORD;
    domain : STRING;
END_VAR

END_FUNCTION

(* ---- DNS_SNTP_SYSLOG_DEMO.st ---- *)
FUNCTION DNS_SNTP_SYSLOG_DEMO
VAR
    IP_C : IP_C;
    S_BUF : NETWORK_BUFFER;
    R_BUF : NETWORK_BUFFER;
    IP_CONTROL_1 : IP_CONTROL;
    DNS_CLIENT : DNS_CLIENT;
    SNTP_CLIENT : SNTP_CLIENT;
    SNTP_SERVER : SNTP_SERVER;
    COUNT_DR : oscat_basic.COUNT_DR;
    RTC_2 : oscat_basic.RTC_2;
    count_cycles : DWORD;
    dns_error : DWORD;
    sntp_error : DWORD;
    freigabe : BOOL;
    dso : BOOL;
    xms : INT;
    sntp_srv_enable : BOOL;
    cur_UDT : DT;
    SYS_LOG : SYS_LOG;
    sys_log_option : BYTE := 2#100;
    TON_1 : TON;
    tp_sys_log : BOOL;
    error_sys_log : DWORD;
    sys_time : TIME;
    cur_LOCAL_DT : DT;
END_VAR

END_FUNCTION

(* ---- DST.st ---- *)
FUNCTION DST : BOOL
VAR_INPUT
    UTC : DT;
END_VAR

VAR
    yr : INT;
    yr4 : DWORD;
    ltc : DWORD;
    idate : DWORD;
END_VAR
yr := YEAR_OF_DATE(DT_TO_DATE(UTC));
ltc := DT_TO_DWORD(UTC);
idate := DT_TO_DWORD(SET_DT(yr, 3, 31, 1, 0, 0));
yr4 := SHR(5 * INT_TO_DWORD(yr), 2) + 1;
DST := (idate - ((yr4 + 3) MOD 7) * 86400 <= ltc) AND (idate + (214 - (yr4) MOD 7) * 86400 > ltc);

(*
Equation used TO calculate the beginning OF European Summer TIME:
Sunday (31 - (5*y/4 + 4) mod 7) March at 01.00 UTC
(valid through 2099, courtesy of Robert H. van Gent, EC).

European Summer Time ends (clocks go back) at 01.00 UTC on

    * 29 October 2006
    * 28 October 2007
    * 26 October 2008

Equation used to calculate the end of European Summer Time:
Sunday (31 - (5*y/4 + 1) mod 7) October at 01.00 UTC
(validity AND credits as above).

*)

(* revision history
hm	4. aug 2006	rev 1.0
	original version

hm	24. okt 2007	rev 1.1
	deleted time_zone_offset input because dst is generally at 01:00 utc and not mesz
	uk starts 01:00 utc and also greece

hm	1. dec 2007	rev 1.2
	changed code to improve performance

hm	16. mar. 2008	rev 1.3
	added type conversion to avoid warnings under codesys 3.0
	code improvement for better performance

hm	7. oct. 2008	rev 1.4
	changed name of function year to year_of_date

hm	24. jan. 2011	rev 1.5
	improved performance
*)
END_FUNCTION

(* ---- DT2_TO_SDT.st ---- *)
FUNCTION DT2_TO_SDT : SDT
VAR_INPUT
    DI : DATE;  // Input variable of type DATE
    TI : TOD;   // Input variable of type TOD
END_VAR
DT2_TO_SDT.YEAR := YEAR_OF_DATE(di);
DT2_TO_SDT.MONTH := MONTH_OF_DATE(di);
DT2_TO_SDT.DAY := DAY_OF_MONTH(di);
DT2_TO_SDT.WEEKDAY := DAY_OF_WEEK(di);
DT2_TO_SDT.MS := DWORD_TO_INT(TOD_TO_DWORD(ti) MOD 1000);
DT2_TO_SDT.SECOND := DWORD_TO_INT((TOD_TO_DWORD(ti) / 1000) MOD 60);
DT2_TO_SDT.MINUTE := DWORD_TO_INT((TOD_TO_DWORD(ti) / 60000) MOD 60);
DT2_TO_SDT.HOUR := DWORD_TO_INT(TOD_TO_DWORD(ti) / 3600000);

(* revision history

hm 18. oct. 2008	rev 1.0
	original version

*)
END_FUNCTION

(* ---- DT_TO_SDT.st ---- *)
FUNCTION DT_TO_SDT : SDT
VAR_INPUT
    DTI : TIME_DT;
END_VAR

VAR
    tmp : DATE;
    tdt : DWORD;
END_VAR
tmp := DT_TO_DATE(dti);
tdt := DT_TO_DWORD(dti) - DATE_TO_DWORD(tmp);
DT_TO_SDT.YEAR := YEAR_OF_DATE(tmp);
DT_TO_SDT.MONTH := MONTH_OF_DATE(tmp);
DT_TO_SDT.DAY := DAY_OF_MONTH(tmp);
DT_TO_SDT.WEEKDAY := DAY_OF_WEEK(tmp);
DT_TO_SDT.SECOND := DWORD_TO_INT(tdt MOD 60);
DT_TO_SDT.MINUTE := DWORD_TO_INT((tdt / 60) MOD 60);
DT_TO_SDT.HOUR := DWORD_TO_INT(tdt / 3600);

(* revision history

hm 18. oct. 2008	rev 1.0
	original version

*)
END_FUNCTION

(* ---- DT_TO_STRF.st ---- *)
FUNCTION DT_TO_STRF : string
VAR_INPUT
    DTI : TIME_DT; // Date and Time Input
    MS : INT;      // Integer Input
    FMT : STRING;  // Format String Input
    LANG : INT;    // Language Input
END_VAR

VAR_CONSTANT
    FILL : STRING[1] := '0'; // Constant String FILL
    BLANK : STRING[1] := ' '; // Constant String BLANK
END_VAR

VAR
    ly : INT;      // Local Integer Variable
    dx : DATE;     // Local Date Variable
    fs : STRING[10]; // Local String Variable (length 10)
    td : TIME_OF_DAY; // Local Time of Day Variable
    tmp : INT;     // Temporary Integer Variable
    pos : INT;     // Position Integer Variable
    f : INT;       // Another Integer Variable
END_VAR
IF LANG < 1 THEN ly := language.DEFAULT; ELSE ly := MIN(language.LMAX, LANG); END_IF;

(* decode date and time information *)
dx := DT_TO_DATE(DTI);
td := DT_TO_TOD(DTI);

(* parse the format string *)
DT_TO_STRF := FMT;
pos := FIND(DT_TO_STRF, '#');
WHILE pos > 0 DO
	(* retrieve format identifier *)
	f := CODE(DT_TO_STRF, pos + 1);
	(* generate the return string according to the format character *)
	fs := '';
	CASE f OF
		65 : (* letter A retunrs the year in 4 digits *)
			fs := INT_TO_STRING(YEAR_OF_DATE(dx));
		66 : (* letter B returns the year in exactly 2 digits *)
			fs := RIGHT(INT_TO_STRING(YEAR_OF_DATE(dx)),2);
		67 : (* letter C returns the month with 1 or 2 digits *)
			fs := INT_TO_STRING(MONTH_OF_DATE(dx));
		68 : (* letter D returns the month with exactly 2 digits *)
			fs := INT_TO_STRING(MONTH_OF_DATE(dx));
			IF LEN(fs) < 2 THEN fs := CONCAT('0', fs); END_IF;
		69 : (* letter E returns the month with 3 characters *)
			fs := MONTH_TO_STRING(MONTH_OF_DATE(dx), ly, 3);
		70 : (* letter F returns the month with all characters *)
			fs := MONTH_TO_STRING(MONTH_OF_DATE(dx), ly, 0);
		71 : (* letter G returns the day with up to 2 digits *)
			fs := INT_TO_STRING(DAY_OF_MONTH(dx));
		72 : (* letter H returns the day of the month with exactly 2 digits *)
			fs := INT_TO_STRING(DAY_OF_MONTH(dx));
			IF LEN(fs) < 2 THEN fs := CONCAT(FILL, fs); END_IF;
		73 : (* letter I returns the weekday as the number 1..7 1 = monday *)
			fs := INT_TO_STRING(DAY_OF_WEEK(dx));
		74 : (* letter J returns the weekday in 2 character writing *)
			fs := WEEKDAY_TO_STRING(DAY_OF_WEEK(dx), ly, 2);
		75 : (* letter K returns the weekday with all characters *)
			fs := WEEKDAY_TO_STRING(DAY_OF_WEEK(dx), ly, 0);
		76 : (* letter L returns AM or PM for the given DateTime *)
			IF td >= TOD#12:00 THEN fs := 'PM'; ELSE fs := 'AM'; END_IF;
		77 : (* letter M returns the hour in 1 or 2 digit form 0..24h *)
			fs := INT_TO_STRING(HOUR(td));
		78 : (* letter N returns the hour in exactly 2 digit form 0..24h *)
			fs := INT_TO_STRING(HOUR(td));
			IF LEN(fs) < 2 THEN fs := CONCAT(FILL, fs); END_IF;
		79 : (* letter O returns the hour in 1 or 2 digit form 0..12h *)
			tmp := HOUR(td) MOD 12;
			IF tmp = 0 THEN tmp := 12; END_IF;
			fs := INT_TO_STRING(tmp);
		80 : (* letter P returns the hour in exactly 2 digit form 0..12h *)
			tmp := HOUR(td) MOD 12;
			IF tmp = 0 THEN tmp := 12; END_IF;
			fs := INT_TO_STRING(tmp);
			IF LEN(fs) < 2 THEN fs := CONCAT(FILL, fs); END_IF;
		81 : (* letter Q returns the minute of the hour in 1 or two digit form *)
			fs := INT_TO_STRING(MINUTE(td));
		82 : (* letter R returns the minute of the hour in exactly two digit form *)
			fs := INT_TO_STRING(MINUTE(td));
			IF LEN(fs) < 2 THEN fs := CONCAT(FILL, fs); END_IF;
		83 : (* letter S returns the second of the minute in 1 or two digit form *)
			fs := INT_TO_STRING(REAL_TO_INT(SECOND(td)));
		84 : (* letter T returns the second of the minute in exactly two digit form *)
			fs := INT_TO_STRING(REAL_TO_INT(SECOND(td)));
			IF LEN(fs) < 2 THEN fs := CONCAT(FILL, fs); END_IF;
		85 : (* letter U returns the milliseconds in 1 to 3 digits *)
			fs := INT_TO_STRING(MS);
		86 : (* letter V returns the milliseconds in exactly 3 digit form *)
			fs := INT_TO_STRING(MS);
			fs := CONCAT('00',fs);
			fs := RIGHT(fs, 3);
		87 : (* letter W returns the day of the month with exactly 2 digits first digit is filled with blank if necessary *)
			fs := INT_TO_STRING(DAY_OF_MONTH(dx));
			IF LEN(fs) < 2 THEN fs := CONCAT(BLANK, fs); END_IF;
		88 : (* letter X returns the month with exactly 2 digits first digit is filled with blank if necessary *)
			fs := INT_TO_STRING(MONTH_OF_DATE(dx));
			IF LEN(fs) < 2 THEN fs := CONCAT(BLANK, fs); END_IF;
		END_CASE;
	DT_TO_STRF := REPLACE(DT_TO_STRF, fs, 2, pos);
	pos := FIND(DT_TO_STRF, '#');
END_WHILE;

(* revision history
hm	7. oct. 2008	rev 1.0
	original version

hm	19. oct. 2008	rev 1.1
	changed language setup constants
*)
END_FUNCTION

(* ---- DW_TO_REAL.st ---- *)
FUNCTION DW_TO_REAL : REAL
VAR_INPUT
    X : DWORD; // Input variable
END_VAR

VAR
    pt : ^REAL; // Pointer to REAL type
END_VAR
pt := ADR(X);
DW_TO_REAL := pt^;

(* revision history
hm	18. apr. 2008
	original version

*)
END_FUNCTION

(* ---- DWORD_OF_BYTE.st ---- *)
FUNCTION DWORD_OF_BYTE : DWORD
VAR_INPUT
    B3 : BYTE;
    B2 : BYTE;
    B1 : BYTE;
    B0 : BYTE;
END_VAR
DWORD_OF_BYTE := SHL(SHL(SHL(BYTE_TO_DWORD(B3),8) OR BYTE_TO_DWORD(B2),8) OR BYTE_TO_DWORD(B1),8) OR BYTE_TO_DWORD(B0);

(* revision history
hm	24. jan 2007	rev 1.0
	original version

hm 2. jan 2008	rev 1.1
	inproved performance

hm	23. apr. 2008	rev 1.2
	reverse order of inputs to be more logical

hm	18. jul. 2009	rev 1.3
	added type conversions for compatibility reasons
*)
END_FUNCTION

(* ---- DWORD_OF_WORD.st ---- *)
FUNCTION DWORD_OF_WORD : DWORD
VAR_INPUT
    W1: WORD;
    W0: WORD;
END_VAR
DWORD_OF_WORD := SHL(WORD_TO_DWORD(W1),16) OR WORD_TO_DWORD(W0);

(* revision history

hm	18. jul. 2009	rev 1.0
	original version

*)
END_FUNCTION

(* ---- DWORD_TO_STRB.st ---- *)
FUNCTION DWORD_TO_STRB : string
VAR_INPUT
    IN : DWORD;
END_VAR_INPUT

VAR
    pt : POINTER TO BYTE;
    i : INT;
END_VAR
(* pointer für die ausgabe ermitteln *)
pt := ADR(DWORD_TO_STRB);
(* die 8 ausgabecharacter ermitteln und schreiben *)
FOR i := 1 TO 32 DO
	pt^:= BOOL_TO_BYTE(in.31) + 48;
	in := SHL(in,1);
	pt := pt + 1;
END_FOR;

(* der ausgabestring muss nochg mit 0 abgeschlossen werden *)
pt^ := 0;

(* revision history
hm		9.6.2007	rev 1.0
	original version

hm		15.dec 2007	rev 1.1
	changed code for better performance

hm	29. mar. 2008	rev 1.2
	changed STRING to STRING(32)

hm	20. jun. 2008	rev 1.3
	performance improvement

*)
END_FUNCTION

(* ---- DWORD_TO_STRF.st ---- *)
FUNCTION DWORD_TO_STRF : string
VAR_INPUT
    IN : DWORD;
    N : INT;
END_VAR
(* limit N to max 20 characters *)
(* convert dword to string first and cut to length N *)
DWORD_TO_STRF := FIX(DWORD_TO_STRING(in),LIMIT(0,N,20),48,1);

(* revision history
hm	26. jan.2007	rev 1.0
	original version

hm	29. mar. 2008	rev 1.1
	changed STRING to STRING(20)
	limit the output string to max 20 digits
*)
END_FUNCTION

(* ---- DWORD_TO_STRH.st ---- *)
FUNCTION DWORD_TO_STRH : string
VAR_INPUT
    IN : DWORD;
END_VAR

VAR
    i : INT;
    temp : BYTE;
    pt : POINTER TO BYTE;
END_VAR
(* read output adress to pointer *)
pt := ADR(DWORD_TO_STRH) + 8;
(* wirte the closing byte for the string *)
pt^:= 0;

(* write the 8 hex characters backwards *)
FOR i := 1 TO 8 DO;
	(* decrement the pointer *)
	pt := pt - 1;
	(* read the lowest order hex value *)
	temp := DWORD_TO_BYTE(in AND 16#0000000F);
	(* convert value to hex character *)
	IF temp <= 9 THEN temp := temp + 48; ELSE temp := temp + 55; END_IF;
	(* write character to output string *)
	PT^ := temp;
	(* shift in for nect hex character *)
	in := SHR(in,4);
END_FOR;

(* code beofre rev 1.2
FOR i := 1 TO 8 DO
	X := DWORD_TO_BYTE(in AND 2#1111);
	IF X <= 9 THEN X := X + 48; ELSE X := X + 55; END_IF;
	Cx := CHR(X);
	temp := CONCAT(Cx, temp);
	in := SHR(in,4);
END_FOR;
DWORD_TO_STRH := temp;
*)

(* revision history
hm	9. jun. 2007	rev 1.0
	original version

hm	11. sep. 2007	rev 1.1
	changed coding for compatibility with twincat, concat cannot support a function as an argument.

hm	15. dec. 2007	rev 1.2
	changed code for better performance

hm	29. mar. 2008	rev 1.3
	changed STRING to STRING(8)

*)
END_FUNCTION

(* ---- EASTER.st ---- *)
FUNCTION EASTER : DATE
VAR_INPUT
    year : INT;
END_VAR

VAR
    b : INT;
    c : INT;
    oday : INT;
END_VAR
b := (204 - 11 * (YEAR MOD 19)) MOD 30;
IF b > 27 THEN b := b - 1; END_IF;
c := (year + SHR(year,2) + b - 13) MOD 7;
oday := 28 + b - c;
IF oday > 33 THEN
	EASTER := SET_DATE(year, 4, oday - 31);
ELSE
	EASTER := SET_DATE(year, 3, oday);
END_IF;

(* alternativer algorithmus ueber das pasah fest
execution time roughly 200us
Der sog. Passah-Vollmond wird berechnet, in dem das Jahr durch 19 ge-
teilt wird und der Rest mit der folgenden Tabelle verglichen wird:

    0: Apr 14       5: Apr 18      10: Mrz 25      15: Mrz 30
    1: Apr 03       6: Apr 08      11: Apr 13      16: Apr 17
    2: Mrz 23       7: Mrz 28      12: Apr 02      17: Apr 07
    3: Apr 11       8: Apr 16      13: Mrz 22      18: Mrz 27
    4: Mrz 31       9: Apr 05      14: Apr 10

Faellt dieses Datum auf einen Sonntag, ist Ostern der naechste Sonntag!

Beispiel: 1992 MOD 19 = 16, daraus folgt 17.04., der naechste Sonntag
          ist dann der 19. April (Ostersonntag)
*)

(* this algorithm is 180 us
a := year MOD 19;
b := year / 100;
c := year MOD 100;
d := b / 4;
e := b MOD 4;
f := (b + 8) / 25;
g := (b - f + 1) / 3;
h := (19 * a + b - d -g + 15) MOD 30;
i := C / 4;
k := c MOD 4;
l := (32 + 2*e + 2*i - h - k) MOD 7;
m := (a + 11 * h + 22 * l) / 451;
x := h + l - 7 * m + 114;
n := X / 31;
o := x MOD 31 + 1;

easter := set_Date(year,n,o);
*)
(*
Im Magazin "Nature" vom 20. April 1876 veröffentlichte ein anonymer Autor eine Tabelle mit Regeln zur Berechnung des (Gregorianischen) Ostersonntages des Jahres J. In Formeln ausgedrückt erhält man das Folgende:
a	=	J mod 19
b	=	int(J / 100)
c	=	J mod 100
d	=	int(b / 4)
e	=	b mod 4
f	=	int((b + 8) / 25)
g	=	int((b - f + 1) / 3
h	=	(19 · a + b - d - g + 15) mod 30
i	=	int(c / 4)
k	=	c mod 4
l	=	(32 + 2 · e + 2 · i - h - k) mod 7
m	=	int((a + 11 · h + 22 · l) / 451)
n	=	int((h + l - 7 · m + 114) / 31)
o	=	(h + l - 7 · m + 114) mod 31

n ist hierbei die Nummer des Monats, o + 1 die Nummer des Tages auf welchen der Ostersonntag im Jahr J fällt. Dieser Algorithmus kommt ohne Hilfszahlen aus.

*)

(* revision history
hm	27. dec 2006	rev 1.0
	original version

hm	15. dec 2007	rev 1.1
	modified code for better performance

hm	3. feb 2008		rev 1.2
	modified code for better performance

hm	7. apr. 2008	rev 1.3
	improved performance
*)
END_FUNCTION

(* ---- ELEMENT_COUNT.st ---- *)
FUNCTION ELEMENT_COUNT : INT
VAR_INPUT
    SEP : BYTE;
END_VAR_INPUT

VAR_IN_OUT
    ELEMENT : STRING[ELEMENT_LENGTH];
END_VAR_IN_OUT

VAR
    pt : POINTER TO ARRAY[1..ELEMENT_LENGTH] OF BYTE;
    l : INT;
    pos : INT;
END_VAR
IF ELEMENT = '' THEN
	ELEMENT_COUNT := 0;
ELSE
	PT := ADR(ELEMENT);
	ELEMENT_COUNT := 1;
	l := LEN(ELEMENT);
	FOR pos := 1 TO l DO
		IF pt^[pos] = SEP THEN ELEMENT_COUNT := ELEMENT_COUNT + 1; END_IF;
	END_FOR;
END_IF;

(* revision histroy
ks	5. apr. 2011	rev 1.0
	original release

*)
END_FUNCTION
